(* IEC 61131-3 sources: guidance-for-physical-ai-production-designer-on-aws/source/plan2cell/examples/welding_cell_2_small/plc/trust/robot1/src, 20 files *)

(* ---- E_PlayerState.st ---- *)
(*
 * E_PlayerState
 * States of FB_ProgramPlayer (robot side of the bt2plc zone protocol).
 * Device simulator R1 (robot1), cell welding_cell_2_small. Generated by bt2plc 0.1.0.
 *)

TYPE E_PlayerState :
(
    PS_IDLE         := 0,    (* No program, pose held *)
    PS_NEXT_OP      := 10,   (* Advance to the next op: wStep := k, REQUEST := mask *)
    PS_WAIT_GRANT   := 20,   (* Wait (GRANT AND mask) = mask *)
    PS_DELAY        := 30,   (* Start delay of the op *)
    PS_MOVE         := 40,   (* Trajectory / blind home move *)
    PS_HOLD         := 50,   (* Hold at the end pose *)
    PS_WAIT_RELEASE := 60,   (* REQUEST := 0, wait (GRANT AND mask) = 0 *)
    PS_DONE         := 90,   (* Program finished *)
    PS_ERROR        := 99    (* Program aborted with an error *)
);
END_TYPE

(* ---- E_ProgramState.st ---- *)
(*
 * E_ProgramState
 * VW VASS standard - robot program states.
 * Device simulator R1 (robot1), cell welding_cell_2_small. Generated by bt2plc 0.1.0.
 *)

TYPE E_ProgramState :
(
    PRG_IDLE     := 0,
    PRG_RUNNING  := 1,
    PRG_STOPPED  := 2,
    PRG_PAUSED   := 3,
    PRG_FINISHED := 4,
    PRG_ERROR    := 5
);
END_TYPE

(* ---- E_RobotMode.st ---- *)
(*
 * E_RobotMode
 * VW VASS standard - KUKA KR C4 robot operating modes.
 * Device simulator R1 (robot1), cell welding_cell_2_small. Generated by bt2plc 0.1.0.
 *)

TYPE E_RobotMode :
(
    MODE_UNKNOWN := 0,
    MODE_T1      := 1,       (* Test mode 1 - reduced speed *)
    MODE_T2      := 2,       (* Test mode 2 - programmed speed *)
    MODE_AUT     := 3,       (* Automatic mode *)
    MODE_EXT     := 4        (* External automatic - PLC controlled *)
);
END_TYPE

(* ---- ST_OpDef.st ---- *)
(*
 * ST_OpDef
 * One op of the bt2plc robot program (row of GVL_Program.aOps).
 * Op k plays waypoints GVL_Program.aWp[nFirstWp..nLastWp] under the zone mask dwZoneMask.
 * Blind home op: bBlindHome = TRUE, nFirstWp = nLastWp = 0 (joint move to arHomeDeg over R_HOME_S).
 * Device simulator R1 (robot1), cell welding_cell_2_small. Generated by bt2plc 0.1.0.
 *)

TYPE ST_OpDef :
STRUCT
    sName           : STRING(32);   (* Operation id, e.g. 'W01' *)
    nFirstWp        : INT;          (* First waypoint index in aWp (0 = none) *)
    nLastWp         : INT;          (* Last waypoint index in aWp (0 = none) *)
    dwZoneMask      : DWORD;        (* REQUEST/GRANT bits (zones 0..30, bit 31 = permit) *)
    tDelay          : TIME;         (* Start delay after the grant *)
    tHold           : TIME;         (* Hold time at the end pose *)
    rDelay_s        : REAL;         (* Start delay in s (used by FB_ProgramPlayer) *)
    rHold_s         : REAL;         (* Hold time in s (used by FB_ProgramPlayer) *)
    rVelScale       : REAL;         (* Velocity scale of the trajectory (1.0 = nominal) *)
    bBlindHome      : BOOL;         (* TRUE = blind joint move to the home pose *)
END_STRUCT
END_TYPE

(* ---- ST_PROFIsafe_Trailer.st ---- *)
(*
 * ST_PROFIsafe_Trailer
 * PROFIsafe trailer - 4 bytes appended by the safety layer (status + 3-byte CRC).
 * Device simulator R1 (robot1), cell welding_cell_2_small. Generated by bt2plc 0.1.0.
 *)

TYPE ST_PROFIsafe_Trailer :
STRUCT
    byStatus        : BYTE;                     (* Status/Control byte *)
    abyCRC          : ARRAY[0..2] OF BYTE;      (* 3-byte CRC *)
END_STRUCT
END_TYPE

(* ---- ST_SafeInput.st ---- *)
(*
 * ST_SafeInput
 * PROFIsafe (Slot 1 - FDIO64) safe inputs: robot -> PLC, 8 bytes user data.
 * GSDML: 8x Unsigned8 Input + F_MessageTrailer4Byte.
 * Device simulator R1 (robot1), cell welding_cell_2_small. Generated by bt2plc 0.1.0.
 *)

TYPE ST_SafeInput :
STRUCT
    (* Byte 0: Safe robot status *)
    bSafe_DrivesOK          : BOOL;   (* Bit 0: Safe drives monitoring OK *)
    bSafe_RobotStopped      : BOOL;   (* Bit 1: Robot safely stopped (SOS/SS1) *)
    bSafe_ReducedSpeed      : BOOL;   (* Bit 2: Safe reduced speed active (SLS) *)
    bSafe_AxisMonitoring    : BOOL;   (* Bit 3: Safe axis range monitoring OK *)
    bSafe_ToolOK            : BOOL;   (* Bit 4: Safe tool monitoring OK *)
    bSafe_WorkspaceOK       : BOOL;   (* Bit 5: Safe workspace monitoring OK *)
    bSafe_Reserved06        : BOOL;   (* Bit 6: Reserved *)
    bSafe_Reserved07        : BOOL;   (* Bit 7: Reserved *)

    (* Byte 1: Safe gate/zone status *)
    bSafe_Gate1Closed       : BOOL;   (* Bit 0: Safety gate 1 closed *)
    bSafe_Gate2Closed       : BOOL;   (* Bit 1: Safety gate 2 closed *)
    bSafe_Gate3Closed       : BOOL;   (* Bit 2: Safety gate 3 closed *)
    bSafe_LightCurtainOK    : BOOL;   (* Bit 3: Light curtain free *)
    bSafe_EStopOK           : BOOL;   (* Bit 4: E-Stop not pressed (NC) *)
    bSafe_EnablingDevice    : BOOL;   (* Bit 5: Enabling device pressed (T1/T2) *)
    bSafe_OperatorSafe      : BOOL;   (* Bit 6: Operator protection OK *)
    bSafe_Reserved17        : BOOL;   (* Bit 7: Reserved *)

    (* Byte 2: Extended safe status *)
    bSafe_STO_Active        : BOOL;   (* Bit 0: Safe Torque Off active *)
    bSafe_SS1_Active        : BOOL;   (* Bit 1: Safe Stop 1 active *)
    bSafe_SS2_Active        : BOOL;   (* Bit 2: Safe Stop 2 active *)
    bSafe_SOS_Active        : BOOL;   (* Bit 3: Safe Operating Stop active *)
    bSafe_SLS_Active        : BOOL;   (* Bit 4: Safely-Limited Speed active *)
    bSafe_SLP_Active        : BOOL;   (* Bit 5: Safely-Limited Position active *)
    bSafe_Reserved26        : BOOL;   (* Bit 6: Reserved *)
    bSafe_FaultPresent      : BOOL;   (* Bit 7: Safety fault present *)

    (* Bytes 3-7: Additional safe signals *)
    bySafe_UserInput3       : BYTE;   (* Byte 3: User safe input *)
    bySafe_UserInput4       : BYTE;   (* Byte 4: User safe input *)
    bySafe_UserInput5       : BYTE;   (* Byte 5: User safe input *)
    bySafe_UserInput6       : BYTE;   (* Byte 6: User safe input *)
    bySafe_UserInput7       : BYTE;   (* Byte 7: User safe input *)
END_STRUCT
END_TYPE

(* ---- ST_SafeOutput.st ---- *)
(*
 * ST_SafeOutput
 * PROFIsafe (Slot 1 - FDIO64) safe outputs: PLC -> robot, 8 bytes user data.
 * GSDML: 8x Unsigned8 Output + F_MessageTrailer4Byte.
 * Device simulator R1 (robot1), cell welding_cell_2_small. Generated by bt2plc 0.1.0.
 *)

TYPE ST_SafeOutput :
STRUCT
    (* Byte 0: Safe control from PLC *)
    bSafe_DriveEnable       : BOOL;   (* Bit 0: Enable drives (safe channel) *)
    bSafe_ExternalEStop     : BOOL;   (* Bit 1: External E-Stop request *)
    bSafe_SafeStop1         : BOOL;   (* Bit 2: Request Safe Stop 1 *)
    bSafe_SafeStop2         : BOOL;   (* Bit 3: Request Safe Stop 2 *)
    bSafe_ReducedSpeedReq   : BOOL;   (* Bit 4: Request safe reduced speed *)
    bSafe_GateOverride      : BOOL;   (* Bit 5: Gate override (maintenance) *)
    bSafe_Reserved06        : BOOL;   (* Bit 6: Reserved *)
    bSafe_Reserved07        : BOOL;   (* Bit 7: Reserved *)

    (* Byte 1: Safe zone control *)
    bSafe_Zone1Enable       : BOOL;   (* Bit 0: Enable workspace zone 1 *)
    bSafe_Zone2Enable       : BOOL;   (* Bit 1: Enable workspace zone 2 *)
    bSafe_Zone3Enable       : BOOL;   (* Bit 2: Enable workspace zone 3 *)
    bSafe_Zone4Enable       : BOOL;   (* Bit 3: Enable workspace zone 4 *)
    bSafe_Reserved14        : BOOL;   (* Bit 4: Reserved *)
    bSafe_Reserved15        : BOOL;   (* Bit 5: Reserved *)
    bSafe_Reserved16        : BOOL;   (* Bit 6: Reserved *)
    bSafe_Reserved17        : BOOL;   (* Bit 7: Reserved *)

    (* Bytes 2-7: Additional safe control *)
    bySafe_UserOutput2      : BYTE;   (* Byte 2: User safe output *)
    bySafe_UserOutput3      : BYTE;   (* Byte 3: User safe output *)
    bySafe_UserOutput4      : BYTE;   (* Byte 4: User safe output *)
    bySafe_UserOutput5      : BYTE;   (* Byte 5: User safe output *)
    bySafe_UserOutput6      : BYTE;   (* Byte 6: User safe output *)
    bySafe_UserOutput7      : BYTE;   (* Byte 7: User safe output *)
END_STRUCT
END_TYPE

(* ---- ST_VASS_ControlWord.st ---- *)
(*
 * ST_VASS_ControlWord
 * VASS PLC control word - output bytes 0-1 (PLC -> robot), Slot 2 DIO256.
 * Device simulator R1 (robot1), cell welding_cell_2_small. Generated by bt2plc 0.1.0.
 *)

TYPE ST_VASS_ControlWord :
STRUCT
    (* Byte 0 *)
    bDrivesOn           : BOOL;   (* Bit 0: Enable drives *)
    bProgStart          : BOOL;   (* Bit 1: Start program *)
    bProgStop           : BOOL;   (* Bit 2: Stop program *)
    bProgCancel         : BOOL;   (* Bit 3: Cancel program *)
    bModeRequest        : BOOL;   (* Bit 4: Request EXT mode *)
    bReset              : BOOL;   (* Bit 5: Reset error *)
    bHomeRequest        : BOOL;   (* Bit 6: Move to home *)
    bConfirm            : BOOL;   (* Bit 7: Confirm/acknowledge *)

    (* Byte 1 *)
    bJobRequest         : BOOL;   (* Bit 8: New job request *)
    bGripperOpen        : BOOL;   (* Bit 9: Open gripper *)
    bGripperClose       : BOOL;   (* Bit 10: Close gripper *)
    bPeriphRelease      : BOOL;   (* Bit 11: Release peripheral *)
    bSpeedOverride      : BOOL;   (* Bit 12: Apply speed override *)
    bReserved13         : BOOL;   (* Bit 13: Reserved *)
    bReserved14         : BOOL;   (* Bit 14: Reserved *)
    bReserved15         : BOOL;   (* Bit 15: Reserved *)
END_STRUCT
END_TYPE

(* ---- ST_VASS_InputTelegram.st ---- *)
(*
 * ST_VASS_InputTelegram
 * Full VASS input telegram - 32 bytes (robot -> PLC), Slot 2 DIO256 inputs.
 * bt2plc use: bytes 4-5 wCurrentStep = op index (GVL_Program.STEP_BYTE),
 *             bytes 16-27 joint angles A1..A6 (FB_JointAngleEncoder),
 *             bytes 28-31 zone REQUEST DWORD LE (GVL_Program.REQ_BYTE).
 * Device simulator R1 (robot1), cell welding_cell_2_small. Generated by bt2plc 0.1.0.
 *)

TYPE ST_VASS_InputTelegram :
STRUCT
    stStatusWord        : ST_VASS_StatusWord;     (* Bytes 0-1:   Status word *)
    wActiveJobNr        : WORD;                   (* Bytes 2-3:   Active job number *)
    wCurrentStep        : WORD;                   (* Bytes 4-5:   Current program step *)
    wSpeedActual        : WORD;                   (* Bytes 6-7:   Actual speed % *)
    wActiveToolNr       : WORD;                   (* Bytes 8-9:   Active tool number *)
    wErrorCode          : WORD;                   (* Bytes 10-11: Active error code *)
    wWarningCode        : WORD;                   (* Bytes 12-13: Active warning code *)
    wPositionX          : INT;                    (* Bytes 14-15: Position X (0.1mm) *)
    wPositionY          : INT;                    (* Bytes 16-17: Position Y (0.1mm) *)
    wPositionZ          : INT;                    (* Bytes 18-19: Position Z (0.1mm) *)
    wUserWord10         : WORD;                   (* Bytes 20-21: User data *)
    wUserWord11         : WORD;                   (* Bytes 22-23: User data *)
    wUserWord12         : WORD;                   (* Bytes 24-25: User data *)
    wUserWord13         : WORD;                   (* Bytes 26-27: User data *)
    wUserWord14         : WORD;                   (* Bytes 28-29: User data *)
    wUserWord15         : WORD;                   (* Bytes 30-31: User data *)
END_STRUCT
END_TYPE

(* ---- ST_VASS_OutputTelegram.st ---- *)
(*
 * ST_VASS_OutputTelegram
 * Full VASS output telegram - 32 bytes (PLC -> robot), Slot 2 DIO256 outputs.
 * bt2plc use: bytes 4-5 PLAN_ID WORD LE during a production job (GVL_Program.PLAN_ID_BYTE),
 *             bytes 12-15 zone GRANT DWORD LE (GVL_Program.GRANT_BYTE).
 * Device simulator R1 (robot1), cell welding_cell_2_small. Generated by bt2plc 0.1.0.
 *)

TYPE ST_VASS_OutputTelegram :
STRUCT
    stControlWord       : ST_VASS_ControlWord;    (* Bytes 0-1:   Control word *)
    wJobNr              : WORD;                   (* Bytes 2-3:   Requested job number *)
    wParameter1         : WORD;                   (* Bytes 4-5:   Parameter 1 *)
    wParameter2         : WORD;                   (* Bytes 6-7:   Parameter 2 *)
    wSpeedOverride      : WORD;                   (* Bytes 8-9:   Speed override % *)
    wToolRequest        : WORD;                   (* Bytes 10-11: Tool change request *)
    wUserWord6          : WORD;                   (* Bytes 12-13: User command data *)
    wUserWord7          : WORD;                   (* Bytes 14-15: User command data *)
    wUserWord8          : WORD;                   (* Bytes 16-17: User command data *)
    wUserWord9          : WORD;                   (* Bytes 18-19: User command data *)
    wUserWord10         : WORD;                   (* Bytes 20-21: User command data *)
    wUserWord11         : WORD;                   (* Bytes 22-23: User command data *)
    wUserWord12         : WORD;                   (* Bytes 24-25: User command data *)
    wUserWord13         : WORD;                   (* Bytes 26-27: User command data *)
    wUserWord14         : WORD;                   (* Bytes 28-29: User command data *)
    wUserWord15         : WORD;                   (* Bytes 30-31: User command data *)
END_STRUCT
END_TYPE

(* ---- ST_VASS_StatusWord.st ---- *)
(*
 * ST_VASS_StatusWord
 * VASS robot status word - input bytes 0-1 (robot -> PLC), Slot 2 DIO256.
 * Device simulator R1 (robot1), cell welding_cell_2_small. Generated by bt2plc 0.1.0.
 *)

TYPE ST_VASS_StatusWord :
STRUCT
    (* Byte 0 *)
    bDrivesPowered      : BOOL;   (* Bit 0: Drives are powered on *)
    bProgRunning        : BOOL;   (* Bit 1: Program is running *)
    bAtHome             : BOOL;   (* Bit 2: Robot at home position *)
    bInPosition         : BOOL;   (* Bit 3: Robot in target position *)
    bModeExt            : BOOL;   (* Bit 4: External automatic mode active *)
    bReady              : BOOL;   (* Bit 5: Robot ready for command *)
    bError              : BOOL;   (* Bit 6: Error present *)
    bWarning            : BOOL;   (* Bit 7: Warning present *)

    (* Byte 1 *)
    bSafetyGateOK       : BOOL;   (* Bit 8: Safety gate closed *)
    bEStopNotActive     : BOOL;   (* Bit 9: E-Stop NOT active (NC logic) *)
    bProgFinished       : BOOL;   (* Bit 10: Program/job finished *)
    bJobAcknowledge     : BOOL;   (* Bit 11: Job number acknowledged *)
    bToolActive         : BOOL;   (* Bit 12: Tool/gripper active *)
    bPartPresent        : BOOL;   (* Bit 13: Part present in gripper *)
    bPeriphReady        : BOOL;   (* Bit 14: Peripheral devices ready *)
    bMaintRequired      : BOOL;   (* Bit 15: Maintenance required *)
END_STRUCT
END_TYPE

(* ---- ST_Waypoint.st ---- *)
(*
 * ST_Waypoint
 * One trajectory waypoint (row of GVL_Program.aWp). Flat fields for portability.
 * rT = seconds from op start; angles in degrees (KUKA A1..A6 after joint sign/offset mapping).
 * Device simulator R1 (robot1), cell welding_cell_2_small. Generated by bt2plc 0.1.0.
 *)

TYPE ST_Waypoint :
STRUCT
    rT              : REAL;         (* Time from op start (s) *)
    rA1             : REAL;         (* Axis 1 (deg) *)
    rA2             : REAL;         (* Axis 2 (deg) *)
    rA3             : REAL;         (* Axis 3 (deg) *)
    rA4             : REAL;         (* Axis 4 (deg) *)
    rA5             : REAL;         (* Axis 5 (deg) *)
    rA6             : REAL;         (* Axis 6 (deg) *)
END_STRUCT
END_TYPE

(* ---- GVL_DeviceParams.st ---- *)
NAMESPACE GVL_DeviceParams
(*
 * GVL_DeviceParams
 * PROFINET device identity parameters.
 * Device simulator R1 (robot1, station kuka-robi1), cell welding_cell_2_small. Generated by bt2plc 0.1.0.
 *
 * These parameters configure how the CODESYS PROFINET Device presents itself
 * on the network. They MUST match what the Siemens PLC expects (from the GSDML).
 *
 * In CODESYS, these are typically set via:
 *   1. The "PROFINET Device IEC Objects" tab in the device editor
 *   2. Or programmatically by writing to the device parameter structure
 *
 * The CODESYS PROFINET Device stack reads these at startup and uses them
 * in DCP responses and during the PROFINET connection establishment.
 *
 * IMPORTANT: The default CODESYS values (VendorId=0x02CC, DeviceId=0x1017)
 * will NOT work with the Siemens PLC that expects KUKA (0x019B / 0x0301).
 * You MUST override them.
 *)

{attribute 'qualified_only'}
VAR_GLOBAL
    (* === KUKA VKRCnexxt Device Identity === *)
    (* These values come from GSDML-V2.25-KUKA-Roboter-GmbH-VKR C4-Device-V1.0 *)

    VENDOR_ID           : UINT        := 16#019B;                 (* KUKA Roboter GmbH *)
    DEVICE_ID           : UINT        := 16#0301;                 (* VKR C4 Device *)
    STATION_TYPE        : STRING(240) := 'KUKA VKR C4';           (* Station type string *)
    DEVICE_TYPE         : STRING(28)  := 'KUKA VKR C4';           (* Device type string *)
    ORDER_ID            : STRING(20)  := 'KUKA VKRC nexxt';       (* Order number *)
    HW_REVISION         : UINT        := 1;                       (* Hardware revision *)
    SW_REV_PREFIX       : USINT       := 16#56;                   (* 'V' in ASCII *)
    SW_REV_MAJOR        : UINT        := 8;                       (* V8.x *)
    SW_REV_MINOR        : UINT        := 2;                       (* x.2 *)
    SW_REV_PATCH        : UINT        := 0;                       (* x.x.0 *)

    (* === Module Identification Numbers (from GSDML) === *)
    MODULE_IDENT_DAP    : DWORD       := DWORD#16#00000301;       (* DAP - Slot 0 *)
    MODULE_IDENT_FDIO64 : DWORD       := DWORD#16#0000008F;       (* PROFIsafe - Slot 1 *)
    MODULE_IDENT_DIO256 : DWORD       := DWORD#16#00001000;       (* VASS telegram - Slot 2 *)
    SUBMODULE_IDENT     : DWORD       := DWORD#16#00000001;       (* Submodule ident (all slots) *)

    (* === PROFIsafe Parameters (Slot 1) === *)
    (* These must match the F-parameter record in the PLC safety configuration *)
    F_SIL_LEVEL         : UINT        := 3;                       (* SIL 3 *)
    F_CRC_LENGTH        : UINT        := 3;                       (* 3-byte CRC *)
    F_WD_TIME_DEFAULT   : UINT        := 500;                     (* Watchdog 500ms *)
    F_BLOCK_ID          : UINT        := 0;                       (* Block ID *)
    F_PAR_CRC_DEFAULT   : UINT        := 16#FF59;                 (* Default F_Par_CRC = 65369 *)
END_VAR
END_NAMESPACE

(* ---- GVL_IO.st ---- *)
NAMESPACE GVL_IO
(*
 * GVL_IO
 * Global variable list for the PROFINET device I/O mapping.
 * Device simulator R1 (robot1, station kuka-robi1), cell welding_cell_2_small. Generated by bt2plc 0.1.0.
 *
 * These variables are mapped to the PROFINET device modules via the I/O Mapping tab.
 * Do NOT use AT addresses - the mapping is done in the device configuration.
 * Only PLC_PRG accesses this GVL: it copies the commands into local images and writes
 * the robot status back as a whole array / as scalars (the FBs never touch GVL_IO).
 *
 * Module mapping (set in I/O Mapping tab of each module):
 *   SafeIO_FDIO64 (Slot 1):
 *     "8 safe digital inputs" channels  -> GVL_IO.bySafeIn0..bySafeIn7
 *     "8 safe digital outputs" channels -> GVL_IO.bySafeOut0..bySafeOut7
 *
 *   VASS_DIO256 (Slot 2):
 *     Input channel  -> GVL_IO.aVassInputData
 *     Output channel -> GVL_IO.aVassOutputData
 *)

{attribute 'qualified_only'}
VAR_GLOBAL
    (* ========================================================================
       SLOT 1 - PROFIsafe FDIO64 Module
       8 individual USINT/BYTE channels per direction
       Map each one to the corresponding "8 safe digital inputs/outputs" row
       ======================================================================== *)

    (* Safe Inputs: Robot -> PLC (mapped to "8 safe digital inputs" channels) *)
    bySafeIn0       : BYTE;     (* Safe input byte 0: Drive status *)
    bySafeIn1       : BYTE;     (* Safe input byte 1: Gate/protection *)
    bySafeIn2       : BYTE;     (* Safe input byte 2: STO/SS1/SS2/SOS/SLS *)
    bySafeIn3       : BYTE;     (* Safe input byte 3: User *)
    bySafeIn4       : BYTE;     (* Safe input byte 4: User *)
    bySafeIn5       : BYTE;     (* Safe input byte 5: User *)
    bySafeIn6       : BYTE;     (* Safe input byte 6: User *)
    bySafeIn7       : BYTE;     (* Safe input byte 7: User *)

    (* Safe Outputs: PLC -> Robot (mapped to "8 safe digital outputs" channels) *)
    bySafeOut0      : BYTE;     (* Safe output byte 0: Drive enable, E-Stop, SS1/SS2 *)
    bySafeOut1      : BYTE;     (* Safe output byte 1: Zone enables *)
    bySafeOut2      : BYTE;     (* Safe output byte 2: User *)
    bySafeOut3      : BYTE;     (* Safe output byte 3: User *)
    bySafeOut4      : BYTE;     (* Safe output byte 4: User *)
    bySafeOut5      : BYTE;     (* Safe output byte 5: User *)
    bySafeOut6      : BYTE;     (* Safe output byte 6: User *)
    bySafeOut7      : BYTE;     (* Safe output byte 7: User *)

    (* ========================================================================
       SLOT 2 - DIO256 VASS Telegram
       32 bytes per direction as arrays
       ======================================================================== *)

    (* VASS Inputs: Robot -> PLC (32 bytes) *)
    aVassInputData      : ARRAY[0..31] OF BYTE;

    (* VASS Outputs: PLC -> Robot (32 bytes) *)
    aVassOutputData     : ARRAY[0..31] OF BYTE;
END_VAR
END_NAMESPACE

(* ---- GVL_Program.st ---- *)
NAMESPACE GVL_Program
(*
 * GVL_Program - generated by bt2plc 0.1.0 - DO NOT EDIT
 * Robot program of robot1 (R1) for plan bt_1790934549_welding_cell_2_small (cell welding_cell_2_small)
 * Angles in degrees (KUKA A1..A6 after joint sign/offset), times in seconds from op start.
 *)
{attribute 'qualified_only'}
VAR_GLOBAL
    (* ========================================================================
       IDENTITY / PROTOCOL
       ======================================================================== *)
    ROBOT_TAG               : STRING(16) := 'R1';
    ROBOT_NS                : STRING(32) := 'robot1';
    ROBOT_INDEX             : WORD := WORD#1;
    PLAN_ID                 : WORD := WORD#16#F77E;             (* must match the head PLC *)
    PROD_FOLGE              : WORD := WORD#11;
    HOME_FOLGE              : WORD := WORD#125;
    JOB_NUMBER_BYTE         : BOOL := FALSE;
    STEP_BYTE               : INT := 4;
    REQ_BYTE                : INT := 28;
    GRANT_BYTE              : INT := 12;
    PLAN_ID_BYTE            : INT := 4;
    R_TASK_S                : REAL := 0.0200;                   (* device MainTask interval *)
    R_HOME_S                : REAL := 7.0000;                   (* blind home duration *)
    R_AT_HOME_TOL_DEG       : REAL := 0.5000;
    R_START_TOL_DEG         : REAL := 1.0000;
    ERR_UNKNOWN_FOLGE       : WORD := WORD#16#0101;
    ERR_PLAN_MISMATCH       : WORD := WORD#16#0103;
    WARN_START_DEVIATION    : WORD := WORD#16#0201;

    (* ========================================================================
       PROGRAM
       ======================================================================== *)
    N_OPS                   : INT := 8;
    N_WP                    : INT := 211;
    arHomeDeg               : ARRAY[1..6] OF REAL := [0.0000, -90.0000, 90.0000, 0.0000, 0.0000, 0.0000];
    aOps                    : ARRAY[1..8] OF ST_OpDef := [
        (sName := 'W01', nFirstWp := 1, nLastWp := 47, dwZoneMask := DWORD#16#00000001, tDelay := T#0MS, tHold := T#500MS, rDelay_s := 0.0000, rHold_s := 0.5000, rVelScale := 1.0000, bBlindHome := FALSE),    (* #1 W01 (weld) *)
        (sName := 'W02', nFirstWp := 48, nLastWp := 68, dwZoneMask := DWORD#16#00000002, tDelay := T#0MS, tHold := T#500MS, rDelay_s := 0.0000, rHold_s := 0.5000, rVelScale := 1.0000, bBlindHome := FALSE),    (* #2 W02 (weld) *)
        (sName := 'W03', nFirstWp := 69, nLastWp := 95, dwZoneMask := DWORD#16#00000001, tDelay := T#0MS, tHold := T#500MS, rDelay_s := 0.0000, rHold_s := 0.5000, rVelScale := 1.0000, bBlindHome := FALSE),    (* #3 W03 (weld) *)
        (sName := 'W06', nFirstWp := 96, nLastWp := 110, dwZoneMask := DWORD#16#00000002, tDelay := T#0MS, tHold := T#500MS, rDelay_s := 0.0000, rHold_s := 0.5000, rVelScale := 1.0000, bBlindHome := FALSE),    (* #4 W06 (weld) *)
        (sName := 'W05', nFirstWp := 111, nLastWp := 137, dwZoneMask := DWORD#16#00000001, tDelay := T#0MS, tHold := T#500MS, rDelay_s := 0.0000, rHold_s := 0.5000, rVelScale := 1.0000, bBlindHome := FALSE),    (* #5 W05 (weld) *)
        (sName := 'W04', nFirstWp := 138, nLastWp := 159, dwZoneMask := DWORD#16#00000002, tDelay := T#0MS, tHold := T#500MS, rDelay_s := 0.0000, rHold_s := 0.5000, rVelScale := 1.0000, bBlindHome := FALSE),    (* #6 W04 (weld) *)
        (sName := 'R1_PARK', nFirstWp := 160, nLastWp := 169, dwZoneMask := DWORD#16#00000001, tDelay := T#0MS, tHold := T#500MS, rDelay_s := 0.0000, rHold_s := 0.5000, rVelScale := 1.0000, bBlindHome := FALSE),    (* #7 R1_PARK (move) *)
        (sName := 'HOME', nFirstWp := 170, nLastWp := 211, dwZoneMask := DWORD#16#00000002, tDelay := T#0MS, tHold := T#0MS, rDelay_s := 0.0000, rHold_s := 0.0000, rVelScale := 1.0000, bBlindHome := FALSE)    (* #8 HOME (home) *)
    ];
    aWp                     : ARRAY[1..211] OF ST_Waypoint := [
        (* op 1 W01 - traj_robot1_W01 *)
        (rT := 0.0000, rA1 := 0.0000, rA2 := -90.0000, rA3 := 90.0000, rA4 := 0.0000, rA5 := 0.0000, rA6 := 0.0000),
        (rT := 0.2677, rA1 := -0.2925, rA2 := -89.9560, rA3 := 90.0355, rA4 := 0.0753, rA5 := 0.1975, rA6 := 0.0896),
        (rT := 0.5350, rA1 := -1.1481, rA2 := -89.8273, rA3 := 90.1392, rA4 := 0.2955, rA5 := 0.7752, rA6 := 0.3515),
        (rT := 0.8027, rA1 := -2.5335, rA2 := -89.6188, rA3 := 90.3072, rA4 := 0.6521, rA5 := 1.7108, rA6 := 0.7756),
        (rT := 1.0703, rA1 := -4.4157, rA2 := -89.3356, rA3 := 90.5354, rA4 := 1.1366, rA5 := 2.9817, rA6 := 1.3518),
        (rT := 1.3377, rA1 := -6.7615, rA2 := -88.9827, rA3 := 90.8198, rA4 := 1.7404, rA5 := 4.5657, rA6 := 2.0699),
        (rT := 1.6053, rA1 := -9.5379, rA2 := -88.5650, rA3 := 91.1564, rA4 := 2.4550, rA5 := 6.4405, rA6 := 2.9199),
        (rT := 1.8730, rA1 := -12.7117, rA2 := -88.0875, rA3 := 91.5412, rA4 := 3.2720, rA5 := 8.5836, rA6 := 3.8915),
        (rT := 2.1403, rA1 := -16.2497, rA2 := -87.5551, rA3 := 91.9702, rA4 := 4.1827, rA5 := 10.9727, rA6 := 4.9746),
        (rT := 2.4080, rA1 := -20.1190, rA2 := -86.9730, rA3 := 92.4393, rA4 := 5.1786, rA5 := 13.5854, rA6 := 6.1591),
        (rT := 2.6757, rA1 := -24.2863, rA2 := -86.3460, rA3 := 92.9446, rA4 := 6.2512, rA5 := 16.3994, rA6 := 7.4349),
        (rT := 2.9430, rA1 := -28.7185, rA2 := -85.6792, rA3 := 93.4820, rA4 := 7.3921, rA5 := 19.3923, rA6 := 8.7918),
        (rT := 3.2107, rA1 := -33.3826, rA2 := -84.9774, rA3 := 94.0475, rA4 := 8.5926, rA5 := 22.5417, rA6 := 10.2196),
        (rT := 3.4783, rA1 := -38.2454, rA2 := -84.2458, rA3 := 94.6371, rA4 := 9.8443, rA5 := 25.8253, rA6 := 11.7083),
        (rT := 3.7457, rA1 := -43.2738, rA2 := -83.4892, rA3 := 95.2467, rA4 := 11.1386, rA5 := 29.2207, rA6 := 13.2477),
        (rT := 4.0133, rA1 := -48.4346, rA2 := -82.7128, rA3 := 95.8725, rA4 := 12.4670, rA5 := 32.7056, rA6 := 14.8276),
        (rT := 4.2810, rA1 := -53.6948, rA2 := -81.9214, rA3 := 96.5102, rA4 := 13.8209, rA5 := 36.2575, rA6 := 16.4379),
        (rT := 4.5483, rA1 := -59.0212, rA2 := -81.1200, rA3 := 97.1561, rA4 := 15.1919, rA5 := 39.8542, rA6 := 18.0685),
        (rT := 4.8160, rA1 := -64.3808, rA2 := -80.3136, rA3 := 97.8059, rA4 := 16.5715, rA5 := 43.4732, rA6 := 19.7093),
        (rT := 5.0837, rA1 := -69.7403, rA2 := -79.5072, rA3 := 98.4557, rA4 := 17.9510, rA5 := 47.0923, rA6 := 21.3500),
        (rT := 5.3510, rA1 := -75.0667, rA2 := -78.7058, rA3 := 99.1015, rA4 := 19.3220, rA5 := 50.6890, rA6 := 22.9806),
        (rT := 5.6187, rA1 := -80.3269, rA2 := -77.9144, rA3 := 99.7393, rA4 := 20.6760, rA5 := 54.2409, rA6 := 24.5910),
        (rT := 5.8863, rA1 := -85.4878, rA2 := -77.1379, rA3 := 100.3650, rA4 := 22.0044, rA5 := 57.7258, rA6 := 26.1709),
        (rT := 6.1537, rA1 := -90.5161, rA2 := -76.3814, rA3 := 100.9747, rA4 := 23.2987, rA5 := 61.1212, rA6 := 27.7103),
        (rT := 6.4213, rA1 := -95.3789, rA2 := -75.6498, rA3 := 101.5643, rA4 := 24.5503, rA5 := 64.4048, rA6 := 29.1989),
        (rT := 6.6890, rA1 := -100.0430, rA2 := -74.9480, rA3 := 102.1298, rA4 := 25.7509, rA5 := 67.5542, rA6 := 30.6268),
        (rT := 6.9563, rA1 := -104.4752, rA2 := -74.2812, rA3 := 102.6671, rA4 := 26.8917, rA5 := 70.5471, rA6 := 31.9836),
        (rT := 7.2240, rA1 := -108.6425, rA2 := -73.6542, rA3 := 103.1724, rA4 := 27.9644, rA5 := 73.3611, rA6 := 33.2594),
        (rT := 7.4917, rA1 := -112.5118, rA2 := -73.0720, rA3 := 103.6415, rA4 := 28.9603, rA5 := 75.9738, rA6 := 34.4439),
        (rT := 7.7590, rA1 := -116.0498, rA2 := -72.5397, rA3 := 104.0705, rA4 := 29.8710, rA5 := 78.3629, rA6 := 35.5271),
        (rT := 8.0267, rA1 := -119.2236, rA2 := -72.0622, rA3 := 104.4553, rA4 := 30.6879, rA5 := 80.5060, rA6 := 36.4987),
        (rT := 8.2943, rA1 := -122.0000, rA2 := -71.6445, rA3 := 104.7919, rA4 := 31.4026, rA5 := 82.3807, rA6 := 37.3486),
        (rT := 8.5617, rA1 := -124.3458, rA2 := -71.2916, rA3 := 105.0764, rA4 := 32.0064, rA5 := 83.9648, rA6 := 38.0668),
        (rT := 8.8293, rA1 := -126.2280, rA2 := -71.0084, rA3 := 105.3046, rA4 := 32.4908, rA5 := 85.2357, rA6 := 38.6430),
        (rT := 9.0970, rA1 := -127.6134, rA2 := -70.7999, rA3 := 105.4725, rA4 := 32.8474, rA5 := 86.1712, rA6 := 39.0671),
        (rT := 9.3643, rA1 := -128.4690, rA2 := -70.6712, rA3 := 105.5763, rA4 := 33.0677, rA5 := 86.7489, rA6 := 39.3290),
        (rT := 9.6320, rA1 := -128.7615, rA2 := -70.6272, rA3 := 105.6117, rA4 := 33.1430, rA5 := 86.9465, rA6 := 39.4186),
        (rT := 9.7320, rA1 := -128.7615, rA2 := -70.2228, rA3 := 105.9156, rA4 := 33.1800, rA5 := 86.8872, rA6 := 39.3731),
        (rT := 9.8320, rA1 := -128.7615, rA2 := -69.6268, rA3 := 106.3586, rA4 := 33.2522, rA5 := 86.7080, rA6 := 39.2426),
        (rT := 9.9320, rA1 := -128.7615, rA2 := -69.3317, rA3 := 106.5670, rA4 := 33.3382, rA5 := 86.3784, rA6 := 39.0108),
        (rT := 10.0320, rA1 := -128.7615, rA2 := -69.0945, rA3 := 106.7257, rA4 := 33.4236, rA5 := 85.9874, rA6 := 38.7386),
        (rT := 10.1320, rA1 := -128.7615, rA2 := -68.8270, rA3 := 106.9027, rA4 := 33.4818, rA5 := 85.6233, rA6 := 38.4888),
        (rT := 10.2320, rA1 := -128.7615, rA2 := -68.5576, rA3 := 107.0760, rA4 := 33.5282, rA5 := 85.2576, rA6 := 38.2401),
        (rT := 10.3320, rA1 := -128.7615, rA2 := -68.2851, rA3 := 107.2465, rA4 := 33.5686, rA5 := 84.8912, rA6 := 37.9919),
        (rT := 10.4320, rA1 := -128.7615, rA2 := -68.0100, rA3 := 107.4140, rA4 := 33.6041, rA5 := 84.5242, rA6 := 37.7441),
        (rT := 10.5320, rA1 := -128.7615, rA2 := -67.6617, rA3 := 107.6183, rA4 := 33.6457, rA5 := 84.0653, rA6 := 37.4348),
        (rT := 10.6320, rA1 := -128.7615, rA2 := -67.4517, rA3 := 107.7396, rA4 := 33.6697, rA5 := 83.7898, rA6 := 37.2493),
        (* op 2 W02 - traj_robot1_W02 *)
        (rT := 0.0000, rA1 := -128.7615, rA2 := -67.4517, rA3 := 107.7396, rA4 := 33.6697, rA5 := 83.7898, rA6 := 37.2493),
        (rT := 0.2820, rA1 := -128.6426, rA2 := -67.6366, rA3 := 107.8186, rA4 := 32.7502, rA5 := 82.9536, rA6 := 37.7433),
        (rT := 0.5643, rA1 := -128.3199, rA2 := -68.1386, rA3 := 108.0329, rA4 := 30.2544, rA5 := 80.6837, rA6 := 39.0840),
        (rT := 0.8463, rA1 := -127.8443, rA2 := -68.8784, rA3 := 108.3488, rA4 := 26.5764, rA5 := 77.3387, rA6 := 41.0597),
        (rT := 1.1283, rA1 := -127.2668, rA2 := -69.7767, rA3 := 108.7324, rA4 := 22.1103, rA5 := 73.2769, rA6 := 43.4588),
        (rT := 1.4103, rA1 := -126.6384, rA2 := -70.7542, rA3 := 109.1498, rA4 := 17.2501, rA5 := 68.8567, rA6 := 46.0696),
        (rT := 1.6927, rA1 := -126.0100, rA2 := -71.7318, rA3 := 109.5672, rA4 := 12.3899, rA5 := 64.4365, rA6 := 48.6804),
        (rT := 1.9747, rA1 := -125.4325, rA2 := -72.6301, rA3 := 109.9508, rA4 := 7.9238, rA5 := 60.3747, rA6 := 51.0796),
        (rT := 2.2567, rA1 := -124.9570, rA2 := -73.3699, rA3 := 110.2667, rA4 := 4.2458, rA5 := 57.0297, rA6 := 53.0553),
        (rT := 2.5390, rA1 := -124.6342, rA2 := -73.8718, rA3 := 110.4810, rA4 := 1.7500, rA5 := 54.7598, rA6 := 54.3960),
        (rT := 2.8210, rA1 := -124.5154, rA2 := -74.0568, rA3 := 110.5600, rA4 := 0.8305, rA5 := 53.9236, rA6 := 54.8899),
        (rT := 2.9210, rA1 := -124.5151, rA2 := -73.6213, rA3 := 110.8768, rA4 := 0.5687, rA5 := 53.3206, rA6 := 55.0767),
        (rT := 3.0210, rA1 := -124.5148, rA2 := -72.9810, rA3 := 111.3378, rA4 := 0.2163, rA5 := 52.4162, rA6 := 55.3282),
        (rT := 3.1210, rA1 := -124.5148, rA2 := -72.6684, rA3 := 111.5513, rA4 := 0.1257, rA5 := 51.9277, rA6 := 55.3932),
        (rT := 3.2210, rA1 := -124.5148, rA2 := -72.4184, rA3 := 111.7128, rA4 := 0.1050, rA5 := 51.5125, rA6 := 55.4084),
        (rT := 3.3210, rA1 := -124.5148, rA2 := -72.1325, rA3 := 111.8956, rA4 := 0.0727, rA5 := 51.0535, rA6 := 55.4318),
        (rT := 3.4210, rA1 := -124.5148, rA2 := -71.8436, rA3 := 112.0754, rA4 := 0.0510, rA5 := 50.5913, rA6 := 55.4476),
        (rT := 3.5210, rA1 := -124.5148, rA2 := -71.5517, rA3 := 112.2520, rA4 := 0.0354, rA5 := 50.1273, rA6 := 55.4590),
        (rT := 3.6210, rA1 := -124.5148, rA2 := -71.2569, rA3 := 112.4255, rA4 := 0.0248, rA5 := 49.6619, rA6 := 55.4668),
        (rT := 3.7210, rA1 := -124.5148, rA2 := -70.8835, rA3 := 112.6373, rA4 := 0.0160, rA5 := 49.0790, rA6 := 55.4732),
        (rT := 3.8210, rA1 := -124.5148, rA2 := -70.6583, rA3 := 112.7632, rA4 := 0.0121, rA5 := 48.7290, rA6 := 55.4761),
        (* op 3 W03 - traj_robot1_W03 *)
        (rT := 0.0000, rA1 := -124.5148, rA2 := -70.6583, rA3 := 112.7632, rA4 := 0.0121, rA5 := 48.7290, rA6 := 55.4761),
        (rT := 0.2767, rA1 := -124.4617, rA2 := -70.7313, rA3 := 112.7862, rA4 := -0.6572, rA5 := 48.6812, rA6 := 55.9965),
        (rT := 0.5530, rA1 := -124.3117, rA2 := -70.9378, rA3 := 112.8512, rA4 := -2.5487, rA5 := 48.5461, rA6 := 57.4671),
        (rT := 0.8297, rA1 := -124.0786, rA2 := -71.2585, rA3 := 112.9524, rA4 := -5.4877, rA5 := 48.3361, rA6 := 59.7523),
        (rT := 1.1063, rA1 := -123.7762, rA2 := -71.6746, rA3 := 113.0835, rA4 := -9.2998, rA5 := 48.0639, rA6 := 62.7161),
        (rT := 1.3830, rA1 := -123.4185, rA2 := -72.1669, rA3 := 113.2386, rA4 := -13.8102, rA5 := 47.7417, rA6 := 66.2230),
        (rT := 1.6593, rA1 := -123.0192, rA2 := -72.7163, rA3 := 113.4118, rA4 := -18.8444, rA5 := 47.3821, rA6 := 70.1371),
        (rT := 1.9360, rA1 := -122.5922, rA2 := -73.3038, rA3 := 113.5970, rA4 := -24.2279, rA5 := 46.9976, rA6 := 74.3228),
        (rT := 2.2127, rA1 := -122.1513, rA2 := -73.9104, rA3 := 113.7882, rA4 := -29.7859, rA5 := 46.6006, rA6 := 78.6441),
        (rT := 2.4893, rA1 := -121.7105, rA2 := -74.5170, rA3 := 113.9794, rA4 := -35.3439, rA5 := 46.2036, rA6 := 82.9655),
        (rT := 2.7657, rA1 := -121.2835, rA2 := -75.1045, rA3 := 114.1646, rA4 := -40.7273, rA5 := 45.8191, rA6 := 87.1511),
        (rT := 3.0423, rA1 := -120.8842, rA2 := -75.6540, rA3 := 114.3378, rA4 := -45.7616, rA5 := 45.4595, rA6 := 91.0652),
        (rT := 3.3190, rA1 := -120.5264, rA2 := -76.1462, rA3 := 114.4929, rA4 := -50.2720, rA5 := 45.1373, rA6 := 94.5721),
        (rT := 3.5953, rA1 := -120.2241, rA2 := -76.5623, rA3 := 114.6241, rA4 := -54.0840, rA5 := 44.8650, rA6 := 97.5360),
        (rT := 3.8720, rA1 := -119.9910, rA2 := -76.8830, rA3 := 114.7252, rA4 := -57.0231, rA5 := 44.6551, rA6 := 99.8211),
        (rT := 4.1487, rA1 := -119.8409, rA2 := -77.0895, rA3 := 114.7902, rA4 := -58.9146, rA5 := 44.5200, rA6 := 101.2917),
        (rT := 4.4253, rA1 := -119.7879, rA2 := -77.1625, rA3 := 114.8133, rA4 := -59.5839, rA5 := 44.4722, rA6 := 101.8121),
        (rT := 4.5377, rA1 := -119.7876, rA2 := -76.7001, rA3 := 115.1416, rA4 := -60.3559, rA5 := 44.3240, rA6 := 102.6809),
        (rT := 4.6505, rA1 := -119.7872, rA2 := -76.0201, rA3 := 115.6192, rA4 := -61.4852, rA5 := 44.0795, rA6 := 103.9753),
        (rT := 4.7505, rA1 := -119.7872, rA2 := -75.6879, rA3 := 115.8405, rA4 := -62.0177, rA5 := 43.8942, rA6 := 104.6450),
        (rT := 4.8505, rA1 := -119.7872, rA2 := -75.4218, rA3 := 116.0082, rA4 := -62.4422, rA5 := 43.7024, rA6 := 105.2177),
        (rT := 4.9505, rA1 := -119.7872, rA2 := -75.1169, rA3 := 116.1984, rA4 := -62.9641, rA5 := 43.4812, rA6 := 105.9117),
        (rT := 5.0505, rA1 := -119.7872, rA2 := -74.8088, rA3 := 116.3854, rA4 := -63.4806, rA5 := 43.2578, rA6 := 106.6047),
        (rT := 5.1505, rA1 := -119.7872, rA2 := -74.4987, rA3 := 116.5684, rA4 := -63.9374, rA5 := 43.0597, rA6 := 107.2204),
        (rT := 5.2505, rA1 := -119.7872, rA2 := -74.1853, rA3 := 116.7483, rA4 := -64.3947, rA5 := 42.8625, rA6 := 107.8387),
        (rT := 5.3505, rA1 := -119.7872, rA2 := -73.7867, rA3 := 116.9688, rA4 := -65.0379, rA5 := 42.5916, rA6 := 108.7077),
        (rT := 5.4505, rA1 := -119.7872, rA2 := -73.5459, rA3 := 117.1000, rA4 := -65.4365, rA5 := 42.4249, rA6 := 109.2463),
        (* op 4 W06 - traj_robot1_W06 *)
        (rT := 0.0000, rA1 := -119.7872, rA2 := -73.5459, rA3 := 117.1000, rA4 := -65.4365, rA5 := 42.4249, rA6 := 109.2463),
        (rT := 0.2930, rA1 := -119.1489, rA2 := -72.8001, rA3 := 114.8711, rA4 := -64.2164, rA5 := 43.4199, rA6 := 108.0229),
        (rT := 0.5860, rA1 := -117.7444, rA2 := -71.1593, rA3 := 109.9675, rA4 := -61.5322, rA5 := 45.6090, rA6 := 105.3312),
        (rT := 0.8790, rA1 := -116.3400, rA2 := -69.5185, rA3 := 105.0638, rA4 := -58.8479, rA5 := 47.7981, rA6 := 102.6395),
        (rT := 1.1720, rA1 := -115.7016, rA2 := -68.7727, rA3 := 102.8349, rA4 := -57.6278, rA5 := 48.7931, rA6 := 101.4160),
        (rT := 1.2720, rA1 := -115.7012, rA2 := -68.3831, rA3 := 103.1319, rA4 := -57.6419, rA5 := 48.7925, rA6 := 101.4570),
        (rT := 1.3720, rA1 := -115.7007, rA2 := -67.8085, rA3 := 103.5655, rA4 := -57.7461, rA5 := 48.7415, rA6 := 101.6606),
        (rT := 1.4720, rA1 := -115.7006, rA2 := -67.5229, rA3 := 103.7711, rA4 := -58.0189, rA5 := 48.5849, rA6 := 102.1462),
        (rT := 1.5720, rA1 := -115.7007, rA2 := -67.2934, rA3 := 103.9284, rA4 := -58.3483, rA5 := 48.3900, rA6 := 102.7163),
        (rT := 1.6720, rA1 := -115.7007, rA2 := -67.0361, rA3 := 104.1022, rA4 := -58.6282, rA5 := 48.2163, rA6 := 103.1755),
        (rT := 1.7720, rA1 := -115.7007, rA2 := -66.7771, rA3 := 104.2724, rA4 := -58.9197, rA5 := 48.0319, rA6 := 103.6366),
        (rT := 1.8720, rA1 := -115.7007, rA2 := -66.5140, rA3 := 104.4406, rA4 := -59.2591, rA5 := 47.8179, rA6 := 104.1645),
        (rT := 1.9720, rA1 := -115.7007, rA2 := -66.2481, rA3 := 104.6058, rA4 := -59.6142, rA5 := 47.5951, rA6 := 104.7081),
        (rT := 2.0720, rA1 := -115.7007, rA2 := -65.9124, rA3 := 104.8068, rA4 := -60.0493, rA5 := 47.3267, rA6 := 105.3635),
        (rT := 2.1720, rA1 := -115.7007, rA2 := -65.7101, rA3 := 104.9261, rA4 := -60.3105, rA5 := 47.1665, rA6 := 105.7542),
        (* op 5 W05 - traj_robot1_W05 *)
        (rT := 0.0000, rA1 := -115.7007, rA2 := -65.7101, rA3 := 104.9261, rA4 := -60.3105, rA5 := 47.1665, rA6 := 105.7542),
        (rT := 0.2757, rA1 := -115.7494, rA2 := -65.7146, rA3 := 104.8564, rA4 := -59.6416, rA5 := 47.2762, rA6 := 105.2455),
        (rT := 0.5517, rA1 := -115.8870, rA2 := -65.7270, rA3 := 104.6592, rA4 := -57.7513, rA5 := 47.5859, rA6 := 103.8079),
        (rT := 0.8273, rA1 := -116.1007, rA2 := -65.7464, rA3 := 104.3529, rA4 := -54.8140, rA5 := 48.0672, rA6 := 101.5740),
        (rT := 1.1030, rA1 := -116.3780, rA2 := -65.7715, rA3 := 103.9556, rA4 := -51.0043, rA5 := 48.6915, rA6 := 98.6766),
        (rT := 1.3787, rA1 := -116.7061, rA2 := -65.8013, rA3 := 103.4855, rA4 := -46.4967, rA5 := 49.4301, rA6 := 95.2484),
        (rT := 1.6547, rA1 := -117.0722, rA2 := -65.8345, rA3 := 102.9609, rA4 := -41.4655, rA5 := 50.2545, rA6 := 91.4221),
        (rT := 1.9303, rA1 := -117.4638, rA2 := -65.8700, rA3 := 102.3998, rA4 := -36.0854, rA5 := 51.1361, rA6 := 87.3303),
        (rT := 2.2060, rA1 := -117.8681, rA2 := -65.9066, rA3 := 101.8205, rA4 := -30.5308, rA5 := 52.0463, rA6 := 83.1058),
        (rT := 2.4820, rA1 := -118.2723, rA2 := -65.9433, rA3 := 101.2413, rA4 := -24.9762, rA5 := 52.9565, rA6 := 78.8814),
        (rT := 2.7577, rA1 := -118.6639, rA2 := -65.9788, rA3 := 100.6802, rA4 := -19.5961, rA5 := 53.8381, rA6 := 74.7896),
        (rT := 3.0333, rA1 := -119.0301, rA2 := -66.0120, rA3 := 100.1555, rA4 := -14.5649, rA5 := 54.6625, rA6 := 70.9633),
        (rT := 3.3093, rA1 := -119.3582, rA2 := -66.0417, rA3 := 99.6854, rA4 := -10.0572, rA5 := 55.4012, rA6 := 67.5351),
        (rT := 3.5850, rA1 := -119.6354, rA2 := -66.0668, rA3 := 99.2881, rA4 := -6.2475, rA5 := 56.0254, rA6 := 64.6377),
        (rT := 3.8607, rA1 := -119.8492, rA2 := -66.0862, rA3 := 98.9818, rA4 := -3.3103, rA5 := 56.5068, rA6 := 62.4038),
        (rT := 4.1363, rA1 := -119.9868, rA2 := -66.0987, rA3 := 98.7847, rA4 := -1.4200, rA5 := 56.8165, rA6 := 60.9662),
        (rT := 4.4123, rA1 := -120.0355, rA2 := -66.1031, rA3 := 98.7149, rA4 := -0.7511, rA5 := 56.9261, rA6 := 60.4575),
        (rT := 4.5123, rA1 := -120.0357, rA2 := -65.7312, rA3 := 99.0104, rA4 := -0.6308, rA5 := 56.7548, rA6 := 60.3791),
        (rT := 4.6123, rA1 := -120.0360, rA2 := -65.1841, rA3 := 99.4405, rA4 := -0.4466, rA5 := 56.4312, rA6 := 60.2589),
        (rT := 4.7123, rA1 := -120.0360, rA2 := -64.9162, rA3 := 99.6405, rA4 := -0.3319, rA5 := 56.0924, rA6 := 60.1840),
        (rT := 4.8123, rA1 := -120.0359, rA2 := -64.7015, rA3 := 99.7923, rA4 := -0.2398, rA5 := 55.7079, rA6 := 60.1236),
        (rT := 4.9123, rA1 := -120.0359, rA2 := -64.4565, rA3 := 99.9636, rA4 := -0.1684, rA5 := 55.2797, rA6 := 60.0766),
        (rT := 5.0123, rA1 := -120.0359, rA2 := -64.2094, rA3 := 100.1316, rA4 := -0.1162, rA5 := 54.8474, rA6 := 60.0420),
        (rT := 5.1123, rA1 := -120.0359, rA2 := -63.9609, rA3 := 100.2959, rA4 := -0.0836, rA5 := 54.4700, rA6 := 60.0204),
        (rT := 5.2123, rA1 := -120.0359, rA2 := -63.7100, rA3 := 100.4571, rA4 := -0.0624, rA5 := 54.0904, rA6 := 60.0063),
        (rT := 5.3123, rA1 := -120.0359, rA2 := -63.3911, rA3 := 100.6546, rA4 := -0.0410, rA5 := 53.5493, rA6 := 59.9919),
        (rT := 5.4123, rA1 := -120.0359, rA2 := -63.1985, rA3 := 100.7720, rA4 := -0.0303, rA5 := 53.2125, rA6 := 59.9847),
        (* op 6 W04 - traj_robot1_W04 *)
        (rT := 0.0000, rA1 := -120.0359, rA2 := -63.1985, rA3 := 100.7720, rA4 := -0.0303, rA5 := 53.2125, rA6 := 59.9847),
        (rT := 0.2773, rA1 := -120.1288, rA2 := -63.1954, rA3 := 100.6111, rA4 := 0.7952, rA5 := 54.0248, rA6 := 59.6456),
        (rT := 0.5547, rA1 := -120.3834, rA2 := -63.1866, rA3 := 100.1699, rA4 := 3.0584, rA5 := 56.2523, rA6 := 58.7158),
        (rT := 0.8317, rA1 := -120.7638, rA2 := -63.1736, rA3 := 99.5107, rA4 := 6.4400, rA5 := 59.5803, rA6 := 57.3266),
        (rT := 1.1090, rA1 := -121.2340, rA2 := -63.1574, rA3 := 98.6957, rA4 := 10.6204, rA5 := 63.6945, rA6 := 55.6092),
        (rT := 1.3863, rA1 := -121.7582, rA2 := -63.1394, rA3 := 97.7873, rA4 := 15.2801, rA5 := 68.2805, rA6 := 53.6950),
        (rT := 1.6637, rA1 := -122.3003, rA2 := -63.1208, rA3 := 96.8478, rA4 := 20.0996, rA5 := 73.0236, rA6 := 51.7151),
        (rT := 1.9407, rA1 := -122.8245, rA2 := -63.1028, rA3 := 95.9394, rA4 := 24.7593, rA5 := 77.6095, rA6 := 49.8008),
        (rT := 2.2180, rA1 := -123.2947, rA2 := -63.0867, rA3 := 95.1245, rA4 := 28.9397, rA5 := 81.7237, rA6 := 48.0834),
        (rT := 2.4953, rA1 := -123.6751, rA2 := -63.0736, rA3 := 94.4653, rA4 := 32.3213, rA5 := 85.0518, rA6 := 46.6942),
        (rT := 2.7727, rA1 := -123.9297, rA2 := -63.0649, rA3 := 94.0240, rA4 := 34.5845, rA5 := 87.2792, rA6 := 45.7644),
        (rT := 3.0500, rA1 := -124.0225, rA2 := -63.0617, rA3 := 93.8631, rA4 := 35.4100, rA5 := 88.0916, rA6 := 45.4253),
        (rT := 3.1500, rA1 := -124.0227, rA2 := -62.7120, rA3 := 94.1541, rA4 := 35.4756, rA5 := 88.0225, rA6 := 45.3131),
        (rT := 3.2500, rA1 := -124.0229, rA2 := -62.1973, rA3 := 94.5779, rA4 := 35.5837, rA5 := 87.8611, rA6 := 45.0952),
        (rT := 3.3500, rA1 := -124.0230, rA2 := -61.9441, rA3 := 94.7757, rA4 := 35.6709, rA5 := 87.6282, rA6 := 44.8479),
        (rT := 3.4500, rA1 := -124.0229, rA2 := -61.7412, rA3 := 94.9258, rA4 := 35.7491, rA5 := 87.3526, rA6 := 44.5802),
        (rT := 3.5500, rA1 := -124.0229, rA2 := -61.5108, rA3 := 95.0942, rA4 := 35.8058, rA5 := 87.0727, rA6 := 44.3314),
        (rT := 3.6500, rA1 := -124.0229, rA2 := -61.2786, rA3 := 95.2593, rA4 := 35.8504, rA5 := 86.7809, rA6 := 44.0868),
        (rT := 3.7500, rA1 := -124.0229, rA2 := -61.0440, rA3 := 95.4214, rA4 := 35.8877, rA5 := 86.4862, rA6 := 43.8484),
        (rT := 3.8500, rA1 := -124.0229, rA2 := -60.8069, rA3 := 95.5807, rA4 := 35.9201, rA5 := 86.1766, rA6 := 43.6056),
        (rT := 3.9500, rA1 := -124.0229, rA2 := -60.5063, rA3 := 95.7751, rA4 := 35.9594, rA5 := 85.7503, rA6 := 43.2784),
        (rT := 4.0500, rA1 := -124.0229, rA2 := -60.3250, rA3 := 95.8907, rA4 := 35.9822, rA5 := 85.4859, rA6 := 43.0775),
        (* op 7 R1_PARK - traj_robot1_R1_PARK *)
        (rT := 0.0000, rA1 := -124.0229, rA2 := -60.3250, rA3 := 95.8907, rA4 := 35.9822, rA5 := 85.4859, rA6 := 43.0775),
        (rT := 0.2863, rA1 := -125.6247, rA2 := -60.4541, rA3 := 95.8014, rA4 := 35.9822, rA5 := 85.4859, rA6 := 43.0775),
        (rT := 0.5727, rA1 := -129.8294, rA2 := -60.7871, rA3 := 95.5713, rA4 := 35.9822, rA5 := 85.4859, rA6 := 43.0775),
        (rT := 0.8590, rA1 := -135.7360, rA2 := -61.2426, rA3 := 95.2570, rA4 := 35.9822, rA5 := 85.4859, rA6 := 43.0775),
        (rT := 1.1453, rA1 := -142.4435, rA2 := -61.7391, rA3 := 94.9151, rA4 := 35.9822, rA5 := 85.4859, rA6 := 43.0775),
        (rT := 1.4317, rA1 := -149.0509, rA2 := -62.1950, rA3 := 94.6020, rA4 := 35.9822, rA5 := 85.4859, rA6 := 43.0775),
        (rT := 1.7180, rA1 := -154.6572, rA2 := -62.5290, rA3 := 94.3745, rA4 := 35.9822, rA5 := 85.4859, rA6 := 43.0775),
        (rT := 2.0047, rA1 := -158.3613, rA2 := -62.6594, rA3 := 94.2891, rA4 := 35.9822, rA5 := 85.4859, rA6 := 43.0775),
        (rT := 2.0880, rA1 := -160.5075, rA2 := -61.5043, rA3 := 95.1253, rA4 := 35.9822, rA5 := 85.4859, rA6 := 43.0775),
        (rT := 2.1713, rA1 := -158.3613, rA2 := -60.3464, rA3 := 95.9536, rA4 := 35.9822, rA5 := 85.4859, rA6 := 43.0775),
        (* op 8 HOME - traj_robot1_n25 *)
        (rT := 0.0000, rA1 := -158.3613, rA2 := -60.3464, rA3 := 95.9536, rA4 := 35.9822, rA5 := 85.4859, rA6 := 43.0775),
        (rT := 0.2032, rA1 := -158.0833, rA2 := -60.3985, rA3 := 95.9432, rA4 := 35.9190, rA5 := 85.3358, rA6 := 43.0018),
        (rT := 0.4062, rA1 := -157.2676, rA2 := -60.5512, rA3 := 95.9125, rA4 := 35.7336, rA5 := 84.8955, rA6 := 42.7800),
        (rT := 0.6095, rA1 := -155.9418, rA2 := -60.7995, rA3 := 95.8626, rA4 := 35.4324, rA5 := 84.1798, rA6 := 42.4193),
        (rT := 0.8127, rA1 := -154.1335, rA2 := -61.1381, rA3 := 95.7947, rA4 := 35.0215, rA5 := 83.2037, rA6 := 41.9274),
        (rT := 1.0160, rA1 := -151.8703, rA2 := -61.5619, rA3 := 95.7096, rA4 := 34.5073, rA5 := 81.9819, rA6 := 41.3118),
        (rT := 1.2190, rA1 := -149.1796, rA2 := -62.0657, rA3 := 95.6084, rA4 := 33.8959, rA5 := 80.5295, rA6 := 40.5799),
        (rT := 1.4222, rA1 := -146.0892, rA2 := -62.6444, rA3 := 95.4922, rA4 := 33.1937, rA5 := 78.8612, rA6 := 39.7392),
        (rT := 1.6255, rA1 := -142.6265, rA2 := -63.2928, rA3 := 95.3621, rA4 := 32.4070, rA5 := 76.9920, rA6 := 38.7973),
        (rT := 1.8288, rA1 := -138.8192, rA2 := -64.0057, rA3 := 95.2189, rA4 := 31.5419, rA5 := 74.9368, rA6 := 37.7616),
        (rT := 2.0317, rA1 := -134.6948, rA2 := -64.7780, rA3 := 95.0639, rA4 := 30.6048, rA5 := 72.7103, rA6 := 36.6397),
        (rT := 2.2350, rA1 := -130.2809, rA2 := -65.6046, rA3 := 94.8979, rA4 := 29.6018, rA5 := 70.3276, rA6 := 35.4390),
        (rT := 2.4382, rA1 := -125.6050, rA2 := -66.4801, rA3 := 94.7221, rA4 := 28.5394, rA5 := 67.8035, rA6 := 34.1671),
        (rT := 2.6415, rA1 := -120.6948, rA2 := -67.3996, rA3 := 94.5375, rA4 := 27.4237, rA5 := 65.1529, rA6 := 32.8314),
        (rT := 2.8445, rA1 := -115.5777, rA2 := -68.3578, rA3 := 94.3452, rA4 := 26.2611, rA5 := 62.3907, rA6 := 31.4395),
        (rT := 3.0478, rA1 := -110.2815, rA2 := -69.3495, rA3 := 94.1460, rA4 := 25.0577, rA5 := 59.5317, rA6 := 29.9988),
        (rT := 3.2510, rA1 := -104.8336, rA2 := -70.3696, rA3 := 93.9412, rA4 := 23.8198, rA5 := 56.5908, rA6 := 28.5168),
        (rT := 3.4542, rA1 := -99.2616, rA2 := -71.4130, rA3 := 93.7317, rA4 := 22.5538, rA5 := 53.5830, rA6 := 27.0012),
        (rT := 3.6572, rA1 := -93.5931, rA2 := -72.4744, rA3 := 93.5186, rA4 := 21.2658, rA5 := 50.5230, rA6 := 25.4592),
        (rT := 3.8605, rA1 := -87.8557, rA2 := -73.5488, rA3 := 93.3029, rA4 := 19.9622, rA5 := 47.4259, rA6 := 23.8985),
        (rT := 4.0637, rA1 := -82.0769, rA2 := -74.6309, rA3 := 93.0857, rA4 := 18.6492, rA5 := 44.3064, rA6 := 22.3266),
        (rT := 4.2668, rA1 := -76.2844, rA2 := -75.7155, rA3 := 92.8679, rA4 := 17.3330, rA5 := 41.1795, rA6 := 20.7509),
        (rT := 4.4700, rA1 := -70.5056, rA2 := -76.7976, rA3 := 92.6507, rA4 := 16.0200, rA5 := 38.0600, rA6 := 19.1789),
        (rT := 4.6732, rA1 := -64.7682, rA2 := -77.8720, rA3 := 92.4350, rA4 := 14.7163, rA5 := 34.9629, rA6 := 17.6183),
        (rT := 4.8765, rA1 := -59.0997, rA2 := -78.9334, rA3 := 92.2219, rA4 := 13.4284, rA5 := 31.9029, rA6 := 16.0763),
        (rT := 5.0795, rA1 := -53.5277, rA2 := -79.9768, rA3 := 92.0124, rA4 := 12.1623, rA5 := 28.8951, rA6 := 14.5606),
        (rT := 5.2828, rA1 := -48.0798, rA2 := -80.9969, rA3 := 91.8076, rA4 := 10.9245, rA5 := 25.9542, rA6 := 13.0787),
        (rT := 5.4860, rA1 := -42.7836, rA2 := -81.9887, rA3 := 91.6085, rA4 := 9.7211, rA5 := 23.0952, rA6 := 11.6380),
        (rT := 5.6892, rA1 := -37.6666, rA2 := -82.9468, rA3 := 91.4161, rA4 := 8.5584, rA5 := 20.3330, rA6 := 10.2461),
        (rT := 5.8922, rA1 := -32.7563, rA2 := -83.8663, rA3 := 91.2315, rA4 := 7.4427, rA5 := 17.6824, rA6 := 8.9104),
        (rT := 6.0955, rA1 := -28.0805, rA2 := -84.7419, rA3 := 91.0557, rA4 := 6.3803, rA5 := 15.1583, rA6 := 7.6385),
        (rT := 6.2987, rA1 := -23.6665, rA2 := -85.5684, rA3 := 90.8897, rA4 := 5.3774, rA5 := 12.7756, rA6 := 6.4378),
        (rT := 6.5020, rA1 := -19.5421, rA2 := -86.3407, rA3 := 90.7347, rA4 := 4.4403, rA5 := 10.5491, rA6 := 5.3159),
        (rT := 6.7050, rA1 := -15.7348, rA2 := -87.0536, rA3 := 90.5916, rA4 := 3.5752, rA5 := 8.4939, rA6 := 4.2802),
        (rT := 6.9082, rA1 := -12.2721, rA2 := -87.7020, rA3 := 90.4614, rA4 := 2.7884, rA5 := 6.6247, rA6 := 3.3383),
        (rT := 7.1115, rA1 := -9.1817, rA2 := -88.2807, rA3 := 90.3452, rA4 := 2.0862, rA5 := 4.9564, rA6 := 2.4976),
        (rT := 7.3147, rA1 := -6.4911, rA2 := -88.7845, rA3 := 90.2440, rA4 := 1.4749, rA5 := 3.5040, rA6 := 1.7657),
        (rT := 7.5177, rA1 := -4.2278, rA2 := -89.2083, rA3 := 90.1589, rA4 := 0.9606, rA5 := 2.2822, rA6 := 1.1500),
        (rT := 7.7210, rA1 := -2.4195, rA2 := -89.5469, rA3 := 90.0910, rA4 := 0.5497, rA5 := 1.3061, rA6 := 0.6582),
        (rT := 7.9242, rA1 := -1.0937, rA2 := -89.7952, rA3 := 90.0411, rA4 := 0.2485, rA5 := 0.5904, rA6 := 0.2975),
        (rT := 8.1273, rA1 := -0.2780, rA2 := -89.9479, rA3 := 90.0105, rA4 := 0.0632, rA5 := 0.1501, rA6 := 0.0756),
        (rT := 8.3305, rA1 := 0.0000, rA2 := -90.0000, rA3 := 90.0000, rA4 := 0.0000, rA5 := 0.0000, rA6 := 0.0000)
    ];
END_VAR
END_NAMESPACE

(* ---- FB_JointAngleEncoder.st ---- *)
(*
 * FB_JointAngleEncoder
 * Device simulator R1 (robot1), cell welding_cell_2_small. Generated by bt2plc 0.1.0.
 *
 * Encodes six KUKA robot joint angles (REAL degrees) into the VASS Option area
 * as scaled fixed-point INTs (0.02 deg per count, big-endian byte order).
 *
 * Encoding per encoding.md:
 *   count = ROUND(angle_deg / 0.02)   clamped to [-32768, +32767]
 *   Byte layout: big-endian (high byte first) in each 2-byte pair
 *
 * Output abyOption = Option area aVassInputData[16..27], 2 bytes per axis
 * (PLC_PRG copies it into the robot -> PLC telegram):
 *   abyOption[0-1]  = bytes 16-17 = A1,  abyOption[2-3]   = bytes 18-19 = A2,
 *   abyOption[4-5]  = bytes 20-21 = A3,  abyOption[6-7]   = bytes 22-23 = A4,
 *   abyOption[8-9]  = bytes 24-25 = A5,  abyOption[10-11] = bytes 26-27 = A6
 *)

FUNCTION_BLOCK FB_JointAngleEncoder
VAR_INPUT
    rA1_deg     : REAL := 0.0;      (* Axis 1 angle in degrees *)
    rA2_deg     : REAL := 0.0;      (* Axis 2 angle in degrees *)
    rA3_deg     : REAL := 0.0;      (* Axis 3 angle in degrees *)
    rA4_deg     : REAL := 0.0;      (* Axis 4 angle in degrees *)
    rA5_deg     : REAL := 0.0;      (* Axis 5 angle in degrees *)
    rA6_deg     : REAL := 0.0;      (* Axis 6 angle in degrees *)
END_VAR

VAR_OUTPUT
    (* Encoded INT values (for monitoring/debug) *)
    iA1_count   : INT;
    iA2_count   : INT;
    iA3_count   : INT;
    iA4_count   : INT;
    iA5_count   : INT;
    iA6_count   : INT;

    (* Option area bytes 16..27 of the robot -> PLC telegram, big-endian A1..A6 *)
    abyOption   : ARRAY[0..11] OF BYTE;
END_VAR

VAR CONSTANT
    SCALE_FACTOR    : REAL := 0.02;     (* degrees per count *)
    INV_SCALE       : REAL := 50.0;     (* 1/0.02 = 50, multiply for speed *)
    COUNT_MAX       : DINT := 32767;
    COUNT_MIN       : DINT := -32768;
END_VAR

VAR
    _arDeg      : ARRAY[1..6] OF REAL;
    _aiCount    : ARRAY[1..6] OF INT;
    _diTemp     : DINT;
    _wTemp      : WORD;
    _i          : INT;
END_VAR
(*
 * FB_JointAngleEncoder - Implementation
 *
 * Converts 6x REAL degree angles to scaled INT counts (0.02 deg per count)
 * and writes them big-endian into abyOption[0..11] (telegram bytes 16..27).
 *
 * Conversion:  count = ROUND(angle / 0.02)  clamped to INT range
 * Byte order:  Big-endian (high byte at lower address) per S7/PROFINET convention
 * Two's complement is formed in DINT (count + 65536 for negative counts), so no
 * bit operation is applied to a signed type.
 *)

_arDeg[1] := rA1_deg;
_arDeg[2] := rA2_deg;
_arDeg[3] := rA3_deg;
_arDeg[4] := rA4_deg;
_arDeg[5] := rA5_deg;
_arDeg[6] := rA6_deg;

FOR _i := 1 TO 6 DO
    (* === Scale and clamp === *)
    _diTemp := REAL_TO_DINT(LIMIT(REAL#-32768.0, _arDeg[_i] * INV_SCALE, REAL#32767.0));
    IF _diTemp > COUNT_MAX THEN _diTemp := COUNT_MAX; END_IF
    IF _diTemp < COUNT_MIN THEN _diTemp := COUNT_MIN; END_IF
    _aiCount[_i] := DINT_TO_INT(_diTemp);

    (* === Big-endian into the Option area: high byte first === *)
    IF _diTemp < 0 THEN
        _diTemp := _diTemp + 65536;
    END_IF
    _wTemp := DINT_TO_WORD(_diTemp);
    abyOption[2 * (_i - 1)] := WORD_TO_BYTE(SHR(_wTemp, 8));
    abyOption[2 * (_i - 1) + 1] := WORD_TO_BYTE(_wTemp AND WORD#16#FF);
END_FOR

iA1_count := _aiCount[1];
iA2_count := _aiCount[2];
iA3_count := _aiCount[3];
iA4_count := _aiCount[4];
iA5_count := _aiCount[5];
iA6_count := _aiCount[6];
END_FUNCTION_BLOCK

(* ---- FB_PROFIsafe_Simulator.st ---- *)
(*
 * FB_PROFIsafe_Simulator
 * Device simulator R1 (robot1), cell welding_cell_2_small. Generated by bt2plc 0.1.0.
 *
 * Simulates the PROFIsafe protocol layer for the FDIO64 module (Slot 1).
 * In a real KUKA controller, the PROFIsafe stack handles CRC generation,
 * sequence counters, and watchdog monitoring.
 *
 * For simulation purposes, this FB:
 * - Monitors the safe output bytes from the PLC (abySafeOut = copy of GVL_IO.bySafeOut0..7)
 * - Provides a "communication OK" flag
 *
 * IMPORTANT: This does NOT provide real functional safety!
 * It only generates data patterns that allow the PLC's PROFIsafe stack
 * to accept the device as communicating. For real safety testing,
 * you need a certified PROFIsafe device or test equipment.
 *
 * PROFIsafe frame structure per IEC 61784-3-3:
 *   [User Data (8 bytes)] [Status/Control (1 byte)] [CRC (3 bytes)]
 *
 * Status byte bits (F_Input from device):
 *   Bit 0: Toggle bit (alternates each cycle)
 *   Bit 1: Reserved
 *   Bit 2: Data valid
 *   Bit 3-7: Reserved / Sequence counter
 *
 * Control byte bits (F_Output from controller):
 *   Bit 0: Toggle bit
 *   Bit 1: Activate device
 *   Bit 2: Reserved
 *   Bit 3-7: Reserved
 *)

FUNCTION_BLOCK FB_PROFIsafe_Simulator
VAR_INPUT
    bEnable         : BOOL := TRUE;
    dwF_Source_Add  : DWORD := DWORD#1;     (* F_Source_Add from parameterization *)
    dwF_Dest_Add    : DWORD := DWORD#1;     (* F_Dest_Add from parameterization *)
    tF_WD_Time      : TIME := T#500MS;      (* Watchdog time *)
    abySafeOut      : ARRAY[0..7] OF BYTE;  (* Safe outputs PLC -> robot (GVL_IO.bySafeOut0..7) *)
END_VAR

VAR_OUTPUT
    bCommOK         : BOOL;                 (* PROFIsafe communication established *)
    bDataValid      : BOOL;                 (* Safe data is valid *)
    bWatchdogError  : BOOL;                 (* Watchdog timeout *)
END_VAR

VAR
    _bToggleBit     : BOOL;                 (* Toggle bit for sequence *)
    _nSeqCounter    : BYTE;                 (* Sequence counter 0-31 *)
    _nCycleCount    : UDINT;                (* Absolute cycle counter *)

    (* Watchdog *)
    _tonWatchdog    : TON;
    _bPLCSafeActive : BOOL;

    (* CRC calculation helper *)
    _dwCrcSeed      : DWORD;
END_VAR
(*
 * FB_PROFIsafe_Simulator - Implementation
 * Works on the input image abySafeOut (PLC_PRG copies GVL_IO.bySafeOut0..7).
 *)

IF NOT bEnable THEN
    bCommOK := FALSE;
    bDataValid := FALSE;
    RETURN;
END_IF

IF _nCycleCount < UDINT#4000000000 THEN
    _nCycleCount := _nCycleCount + 1;
ELSE
    _nCycleCount := 0;
END_IF

(* ============================================================================
   MONITOR PLC SAFE OUTPUT DATA
   ============================================================================ *)
_bPLCSafeActive := (abySafeOut[0] <> BYTE#0) OR (abySafeOut[1] <> BYTE#0);

(* Watchdog *)
_tonWatchdog(IN := NOT _bPLCSafeActive, PT := tF_WD_Time);
bWatchdogError := _tonWatchdog.Q;

bCommOK := _bPLCSafeActive AND NOT bWatchdogError;
bDataValid := bCommOK;
END_FUNCTION_BLOCK

(* ---- FB_ProgramPlayer.st ---- *)
(*
 * FB_ProgramPlayer
 * Device simulator R1 (robot1), cell welding_cell_2_small, tree bt_1790934549_welding_cell_2_small. Generated by bt2plc 0.1.0.
 *
 * Plays the bt2plc robot program (GVL_Program) for PROD_FOLGE, or a blind joint
 * move to the home pose for HOME_FOLGE. Robot side of the zone protocol, per op k
 * with mask M = GVL_Program.aOps[k].dwZoneMask:
 *   1  wStep := k                          (also for M = 0)
 *   2  if M <> 0: REQUEST := M             (same call / telegram as wStep)
 *   3  if M <> 0: wait (GRANT AND M) = M
 *   4  start delay; trajectory (x rVelScale x override); hold
 *   5  if M <> 0: REQUEST := 0
 *   6  if M <> 0: wait (GRANT AND M) = 0   (4-phase, before the next REQUEST)
 *   7  next op; after the last op: bDone, wStep := 0 (same call)
 *
 * Timing: all times are REAL seconds accumulated from rDt (seconds per call, the
 * device task interval). Motion time advances by rDt * rRate * rVelScale, delay and
 * hold by rDt (the override does not scale dwell times). No TIME() / TON is used.
 * Zero-time transitions fall through within one call (at most N_MAX_TRANSITIONS),
 * but wStep changes at most once per call, so every step is visible to the head PLC.
 * Joints (deg) are linearly interpolated between waypoints and published as rA1..rA6_deg.
 * Abort (bAbort level while busy): REQUEST := 0, wStep := 0, the pose is held.
 * The robot powers up at GVL_Program.arHomeDeg.
 *)

FUNCTION_BLOCK FB_ProgramPlayer
VAR_INPUT
    bStart          : BOOL;                 (* Rising edge: start wJob *)
    wJob            : WORD;                 (* Folge to play: PROD_FOLGE or HOME_FOLGE *)
    bAbort          : BOOL;                 (* Level: stop / cancel / drives off / E-stop *)
    dwGrant         : DWORD;                (* Zone GRANT bits from the head PLC *)
    rRate           : REAL := 1.0;          (* Speed override factor (1.0 = 100 %) *)
    rDt             : REAL := 0.02;         (* Seconds per call (task interval) *)
END_VAR

VAR_OUTPUT
    eState          : E_PlayerState;        (* Current state *)
    bBusy           : BOOL;                 (* Program running *)
    bDone           : BOOL;                 (* Latched until next start *)
    bError          : BOOL;                 (* Latched until next start *)
    wErrorCode      : WORD;                 (* Error code, GVL_Program.ERR_xxx *)
    wWarningCode    : WORD;                 (* Warning code, GVL_Program.WARN_xxx, latched until next start *)
    wStep           : WORD;                 (* 1-based op index, 0 = none *)
    dwRequest       : DWORD;                (* Zone REQUEST bits to the head PLC *)
    bAtHome         : BOOL;                 (* All joints within R_AT_HOME_TOL_DEG of arHomeDeg *)
    rA1_deg         : REAL;                 (* Axis 1 angle *)
    rA2_deg         : REAL;                 (* Axis 2 angle *)
    rA3_deg         : REAL;                 (* Axis 3 angle *)
    rA4_deg         : REAL;                 (* Axis 4 angle *)
    rA5_deg         : REAL;                 (* Axis 5 angle *)
    rA6_deg         : REAL;                 (* Axis 6 angle *)
END_VAR

VAR CONSTANT
    N_MAX_TRANSITIONS : INT := 8;           (* Fall-through bound per call *)
END_VAR

VAR
    _eState         : E_PlayerState := E_PlayerState#PS_IDLE;
    _rtrigStart     : R_TRIG;
    _bFirstCall     : BOOL := TRUE;

    (* === Current op === *)
    _nOp            : INT;                  (* 1-based op index, 0 = HOME_FOLGE move *)
    _dwMask         : DWORD;                (* Zone mask of the current op *)
    _bHomeMove      : BOOL;                 (* Current move is a blind home move *)
    _nWp            : INT;                  (* Current waypoint segment start *)
    _nLast          : INT;                  (* Last waypoint of the current op, 0 = none *)
    _rVel           : REAL;                 (* Velocity scale of the current move *)

    (* === Time (s) === *)
    _rDtCall        : REAL;                 (* rDt limited to 0..1 s *)
    _rRateCall      : REAL;                 (* rRate limited to >= 0 *)
    _rT             : REAL;                 (* Motion time since move start *)
    _rTimer         : REAL;                 (* Delay / hold timer *)
    _rDur           : REAL;                 (* Duration of the blind home move *)
    _rAlpha         : REAL;                 (* Interpolation factor 0..1 *)
    _rSpan          : REAL;                 (* Waypoint segment duration *)

    (* === Pose (deg) === *)
    _arQ            : ARRAY[1..6] OF REAL;  (* Current joint angles *)
    _arQ0           : ARRAY[1..6] OF REAL;  (* Pose at the start of a blind home move *)
    _arQa           : ARRAY[1..6] OF REAL;  (* Segment start waypoint *)
    _arQb           : ARRAY[1..6] OF REAL;  (* Segment end waypoint *)

    (* === Fall-through === *)
    _nPass          : INT;
    _bAdvance       : BOOL;                 (* A transition happened in this pass *)
    _bStepSet       : BOOL;                 (* wStep changed in this call *)
    _bMoveDone      : BOOL;
    _i              : INT;
END_VAR
(*
 * FB_ProgramPlayer - Implementation
 *)

(* ============================================================================
   INIT - the robot powers up at the home pose
   ============================================================================ *)
IF _bFirstCall THEN
    FOR _i := 1 TO 6 DO
        _arQ[_i] := GVL_Program.arHomeDeg[_i];
    END_FOR
    _bFirstCall := FALSE;
END_IF

_rDtCall := LIMIT(0.0, rDt, 1.0);
_rRateCall := MAX(rRate, 0.0);
_rtrigStart(CLK := bStart);

(* ============================================================================
   ABORT - stop / cancel / drives off / E-stop: REQUEST := 0, wStep := 0, hold pose
   ============================================================================ *)
IF bAbort AND bBusy THEN
    _eState := E_PlayerState#PS_IDLE;
    bBusy := FALSE;
    wStep := WORD#0;
    dwRequest := DWORD#0;
END_IF

(* ============================================================================
   CLOCK - advance the timer of the state that is active at the start of the call
   (a state entered during this call starts counting with the next call)
   ============================================================================ *)
IF _eState = E_PlayerState#PS_DELAY OR _eState = E_PlayerState#PS_HOLD THEN
    _rTimer := _rTimer + _rDtCall;
ELSIF _eState = E_PlayerState#PS_MOVE THEN
    _rT := _rT + _rDtCall * _rRateCall * _rVel;
END_IF

(* ============================================================================
   START
   ============================================================================ *)
IF _rtrigStart.Q AND NOT bBusy AND NOT bAbort THEN
    bDone := FALSE;
    bError := FALSE;
    wErrorCode := WORD#0;
    wWarningCode := WORD#0;
    wStep := WORD#0;
    dwRequest := DWORD#0;
    _nOp := 0;
    _dwMask := DWORD#0;
    _rT := 0.0;
    _rTimer := 0.0;
    IF wJob = GVL_Program.HOME_FOLGE THEN
        (* Blind joint move from the current pose to arHomeDeg: no step, no zones *)
        FOR _i := 1 TO 6 DO
            _arQ0[_i] := _arQ[_i];
        END_FOR
        _bHomeMove := TRUE;
        _nLast := 0;
        _rVel := 1.0;
        _rDur := GVL_Program.R_HOME_S;
        bBusy := TRUE;
        _eState := E_PlayerState#PS_MOVE;
    ELSIF wJob = GVL_Program.PROD_FOLGE AND GVL_Program.N_OPS > 0 THEN
        bBusy := TRUE;
        _eState := E_PlayerState#PS_NEXT_OP;
    ELSE
        wErrorCode := GVL_Program.ERR_UNKNOWN_FOLGE;
        _eState := E_PlayerState#PS_ERROR;
    END_IF
END_IF

(* ============================================================================
   STATE MACHINE - falls through zero-time transitions (bounded)
   ============================================================================ *)
_bStepSet := FALSE;
FOR _nPass := 1 TO N_MAX_TRANSITIONS DO
    _bAdvance := FALSE;

    CASE _eState OF

    E_PlayerState#PS_IDLE:
        bBusy := FALSE;
        wStep := WORD#0;
        dwRequest := DWORD#0;

    E_PlayerState#PS_NEXT_OP:
        (* wStep changes at most once per call: the head checks step + 1 per telegram *)
        IF NOT _bStepSet THEN
            _nOp := _nOp + 1;
            IF _nOp > GVL_Program.N_OPS THEN
                _eState := E_PlayerState#PS_DONE;
            ELSE
                wStep := INT_TO_WORD(_nOp);
                _bStepSet := TRUE;
                _dwMask := GVL_Program.aOps[_nOp].dwZoneMask;
                IF _dwMask <> DWORD#0 THEN
                    dwRequest := _dwMask;           (* same telegram as wStep *)
                    _eState := E_PlayerState#PS_WAIT_GRANT;
                ELSE
                    _rTimer := 0.0;
                    _eState := E_PlayerState#PS_DELAY;
                END_IF
            END_IF
            _bAdvance := TRUE;
        END_IF

    E_PlayerState#PS_WAIT_GRANT:
        IF (dwGrant AND _dwMask) = _dwMask THEN
            _rTimer := 0.0;
            _eState := E_PlayerState#PS_DELAY;
            _bAdvance := TRUE;
        END_IF

    E_PlayerState#PS_DELAY:
        IF _rTimer >= GVL_Program.aOps[_nOp].rDelay_s THEN
            (* Begin the motion of op _nOp *)
            _rT := 0.0;
            _rVel := GVL_Program.aOps[_nOp].rVelScale;
            IF _rVel <= 0.0 THEN
                _rVel := 1.0;
            END_IF
            _bHomeMove := GVL_Program.aOps[_nOp].bBlindHome;
            IF _bHomeMove THEN
                FOR _i := 1 TO 6 DO
                    _arQ0[_i] := _arQ[_i];
                END_FOR
                _rDur := GVL_Program.R_HOME_S;
                _nLast := 0;
            ELSE
                _nWp := GVL_Program.aOps[_nOp].nFirstWp;
                _nLast := GVL_Program.aOps[_nOp].nLastWp;
                IF _nWp < 1 OR _nLast < _nWp OR _nLast > GVL_Program.N_WP THEN
                    _nLast := 0;                    (* no valid trajectory: zero-length move *)
                ELSE
                    (* Start deviation: the trajectory should start at the current pose *)
                    _arQa[1] := GVL_Program.aWp[_nWp].rA1;
                    _arQa[2] := GVL_Program.aWp[_nWp].rA2;
                    _arQa[3] := GVL_Program.aWp[_nWp].rA3;
                    _arQa[4] := GVL_Program.aWp[_nWp].rA4;
                    _arQa[5] := GVL_Program.aWp[_nWp].rA5;
                    _arQa[6] := GVL_Program.aWp[_nWp].rA6;
                    FOR _i := 1 TO 6 DO
                        IF ABS(_arQ[_i] - _arQa[_i]) > GVL_Program.R_START_TOL_DEG THEN
                            wWarningCode := GVL_Program.WARN_START_DEVIATION;
                        END_IF
                    END_FOR
                END_IF
            END_IF
            _eState := E_PlayerState#PS_MOVE;
            _bAdvance := TRUE;
        END_IF

    E_PlayerState#PS_MOVE:
        _bMoveDone := FALSE;
        IF _bHomeMove THEN
            (* Blind joint move: linear in joint space over R_HOME_S *)
            IF _rDur > 0.0 THEN
                _rAlpha := LIMIT(0.0, _rT / _rDur, 1.0);
            ELSE
                _rAlpha := 1.0;
            END_IF
            FOR _i := 1 TO 6 DO
                _arQ[_i] := _arQ0[_i] + _rAlpha * (GVL_Program.arHomeDeg[_i] - _arQ0[_i]);
            END_FOR
            _bMoveDone := _rAlpha >= 1.0;
        ELSIF _nLast < 1 THEN
            _bMoveDone := TRUE;
        ELSE
            (* Trajectory: find the segment [_nWp, _nWp + 1] that contains _rT *)
            WHILE _nWp < _nLast DO
                IF GVL_Program.aWp[_nWp + 1].rT <= _rT THEN
                    _nWp := _nWp + 1;
                ELSE
                    EXIT;
                END_IF
            END_WHILE
            _arQa[1] := GVL_Program.aWp[_nWp].rA1;
            _arQa[2] := GVL_Program.aWp[_nWp].rA2;
            _arQa[3] := GVL_Program.aWp[_nWp].rA3;
            _arQa[4] := GVL_Program.aWp[_nWp].rA4;
            _arQa[5] := GVL_Program.aWp[_nWp].rA5;
            _arQa[6] := GVL_Program.aWp[_nWp].rA6;
            IF _nWp >= _nLast THEN
                FOR _i := 1 TO 6 DO
                    _arQ[_i] := _arQa[_i];
                END_FOR
                _bMoveDone := TRUE;
            ELSE
                _arQb[1] := GVL_Program.aWp[_nWp + 1].rA1;
                _arQb[2] := GVL_Program.aWp[_nWp + 1].rA2;
                _arQb[3] := GVL_Program.aWp[_nWp + 1].rA3;
                _arQb[4] := GVL_Program.aWp[_nWp + 1].rA4;
                _arQb[5] := GVL_Program.aWp[_nWp + 1].rA5;
                _arQb[6] := GVL_Program.aWp[_nWp + 1].rA6;
                _rSpan := GVL_Program.aWp[_nWp + 1].rT - GVL_Program.aWp[_nWp].rT;
                IF _rSpan > 0.0 THEN
                    _rAlpha := LIMIT(0.0, (_rT - GVL_Program.aWp[_nWp].rT) / _rSpan, 1.0);
                ELSE
                    _rAlpha := 1.0;
                END_IF
                FOR _i := 1 TO 6 DO
                    _arQ[_i] := _arQa[_i] + _rAlpha * (_arQb[_i] - _arQa[_i]);
                END_FOR
            END_IF
        END_IF
        IF _bMoveDone THEN
            IF _nOp = 0 THEN
                _eState := E_PlayerState#PS_DONE;   (* HOME_FOLGE finished *)
            ELSE
                _rTimer := 0.0;
                _eState := E_PlayerState#PS_HOLD;
            END_IF
            _bAdvance := TRUE;
        END_IF

    E_PlayerState#PS_HOLD:
        IF _rTimer >= GVL_Program.aOps[_nOp].rHold_s THEN
            IF _dwMask <> DWORD#0 THEN
                dwRequest := DWORD#0;
                _eState := E_PlayerState#PS_WAIT_RELEASE;
            ELSE
                _eState := E_PlayerState#PS_NEXT_OP;
            END_IF
            _bAdvance := TRUE;
        END_IF

    E_PlayerState#PS_WAIT_RELEASE:
        (* 4-phase: the GRANT must drop before the next REQUEST *)
        IF (dwGrant AND _dwMask) = DWORD#0 THEN
            _eState := E_PlayerState#PS_NEXT_OP;
            _bAdvance := TRUE;
        END_IF

    E_PlayerState#PS_DONE:
        bBusy := FALSE;
        bDone := TRUE;
        wStep := WORD#0;
        dwRequest := DWORD#0;
        _eState := E_PlayerState#PS_IDLE;

    E_PlayerState#PS_ERROR:
        bBusy := FALSE;
        bError := TRUE;
        wStep := WORD#0;
        dwRequest := DWORD#0;
        _eState := E_PlayerState#PS_IDLE;

    END_CASE

    IF NOT _bAdvance THEN
        EXIT;
    END_IF
END_FOR

(* ============================================================================
   PUBLISH
   ============================================================================ *)
bAtHome := TRUE;
FOR _i := 1 TO 6 DO
    IF ABS(_arQ[_i] - GVL_Program.arHomeDeg[_i]) > GVL_Program.R_AT_HOME_TOL_DEG THEN
        bAtHome := FALSE;
    END_IF
END_FOR
rA1_deg := _arQ[1];
rA2_deg := _arQ[2];
rA3_deg := _arQ[3];
rA4_deg := _arQ[4];
rA5_deg := _arQ[5];
rA6_deg := _arQ[6];
eState := _eState;
END_FUNCTION_BLOCK

(* ---- FB_VASS_DeviceSimulator.st ---- *)
(*
 * FB_VASS_DeviceSimulator
 * Device simulator R1 (robot1, station kuka-robi1), cell welding_cell_2_small, tree bt_1790934549_welding_cell_2_small.
 * Generated by bt2plc 0.1.0.
 *
 * Simulates a KUKA KR C4 robot responding to VW VASS commands via PROFINET.
 *
 * This FB reads the PLC commands from its input images (PLC -> robot):
 *   aVassOutputData = copy of GVL_IO.aVassOutputData, abySafeOut = GVL_IO.bySafeOut0..7
 * and produces the robot status images (robot -> PLC):
 *   aVassInputData (bytes 16-27 = 0, the joint encoder fills them in PLC_PRG), abySafeIn.
 * PLC_PRG copies the images from / to GVL_IO; this FB never accesses GVL_IO.
 *
 * Job handshake (as the original simulator): drives on after 2 s, EXT mode, Ready,
 * JobRequest edge -> JobAck + job echo (clears ProgFinished), ProgStart edge -> start,
 * Stop/Cancel level -> stop, Reset held 500 ms -> clear error, gripper, speed override.
 * Job execution is delegated to FB_ProgramPlayer (GVL_Program):
 *   PROD_FOLGE: the bt2plc program; PLAN_ID (bytes PLAN_ID_BYTE..+1, latched at job accept)
 *               must equal GVL_Program.PLAN_ID at ProgStart, else ERR_PLAN_MISMATCH, no start.
 *   HOME_FOLGE: blind joint move to arHomeDeg (also on a HomeRequest [0].6 edge while Ready).
 *   other:      ERR_UNKNOWN_FOLGE, no start.
 * Zone protocol: wCurrentStep at bytes STEP_BYTE..+1, REQUEST DWORD LE at REQ_BYTE..+3,
 * GRANT DWORD LE read from bytes GRANT_BYTE..+3 (GVL_Program offsets).
 * At the end ProgRunning := FALSE, ProgFinished := TRUE and step := 0 in the same scan.
 *)

FUNCTION_BLOCK FB_VASS_DeviceSimulator
VAR_INPUT
    bEnable             : BOOL := TRUE;             (* Enable simulation *)
    wRobotID            : WORD := WORD#1;           (* Robot identification number 1-8 *)
    aVassOutputData     : ARRAY[0..31] OF BYTE;     (* VASS telegram PLC -> robot (GVL_IO.aVassOutputData) *)
    abySafeOut          : ARRAY[0..7] OF BYTE;      (* Safe outputs PLC -> robot (GVL_IO.bySafeOut0..7) *)
    rDt                 : REAL := 0.02;             (* Task interval in s (GVL_Program.R_TASK_S) *)
END_VAR

VAR_OUTPUT
    bActive             : BOOL;                     (* Simulator is active *)
    eCurrentMode        : E_RobotMode;              (* Current operating mode *)
    eProgramState       : E_ProgramState;           (* Current program state *)
    bSafetyOK           : BOOL;                     (* Safety system healthy *)
    aVassInputData      : ARRAY[0..31] OF BYTE;     (* VASS telegram robot -> PLC (bytes 16-27 = 0) *)
    abySafeIn           : ARRAY[0..7] OF BYTE;      (* Safe inputs robot -> PLC (GVL_IO.bySafeIn0..7) *)

    (* Joint angles from the program player (deg) *)
    rA1_deg             : REAL;
    rA2_deg             : REAL;
    rA3_deg             : REAL;
    rA4_deg             : REAL;
    rA5_deg             : REAL;
    rA6_deg             : REAL;

    (* Diagnostics *)
    wActiveJob          : WORD;                     (* Accepted job number (Folge) *)
    wCurrentStep        : WORD;                     (* Current op index, 0 = none *)
    wErrorCode          : WORD;                     (* Active error code *)
    dwRequest           : DWORD;                    (* Zone REQUEST bits sent to the head PLC *)
    dwGrant             : DWORD;                    (* Zone GRANT bits received from the head PLC *)
    ePlayerState        : E_PlayerState;            (* State of the program player *)
END_VAR

VAR
    (* === Internal Robot State === *)
    _bDrivesPowered     : BOOL;
    _bInExtMode         : BOOL;
    _bReady             : BOOL;
    _bError             : BOOL;
    _bProgRunning       : BOOL;
    _bAtHome            : BOOL := TRUE;
    _bInPosition        : BOOL := TRUE;
    _bProgFinished      : BOOL;
    _bJobAcknowledged   : BOOL;
    _bGripperClosed     : BOOL;
    _bPartPresent       : BOOL;
    _bPeriphReady       : BOOL := TRUE;

    _wActiveJob         : WORD;
    _wCurrentStep       : WORD;
    _wSpeed             : WORD := WORD#100;
    _wToolNr            : WORD := WORD#1;
    _wErrorCode         : WORD;
    _wWarningCode       : WORD;

    (* Simulated position (0.1mm units) *)
    _iPositionX         : INT := 5000;              (* 500.0 mm *)
    _iPositionY         : INT := 0;
    _iPositionZ         : INT := 10000;             (* 1000.0 mm *)

    (* === Safety State === *)
    _bSafe_DrivesOK     : BOOL := TRUE;
    _bSafe_Stopped      : BOOL := TRUE;
    _bSafe_EStopOK      : BOOL := TRUE;
    _bSafe_GatesClosed  : BOOL := TRUE;
    _bSafe_Fault        : BOOL;
    _bSafe_STO          : BOOL;
    _bSafe_SS1          : BOOL;

    (* PROFIsafe CRC simulation *)
    _bySafeTrailerStatus : BYTE;
    _nSafeCycleCount     : UDINT;

    (* === Timers === *)
    _tonDriveStartup    : TON;                      (* Simulate drive power-on delay *)
    _tonErrorReset      : TON;                      (* Simulate error reset delay *)
    _tonGripperAction   : TON;                      (* Simulate gripper open/close time *)

    (* === Edge Detection === *)
    _rtrigProgStart     : R_TRIG;
    _rtrigProgStop      : R_TRIG;
    _rtrigReset         : R_TRIG;
    _rtrigJobReq        : R_TRIG;
    _rtrigDrivesOn      : R_TRIG;
    _rtrigHome          : R_TRIG;
    _rtrigGripOpen      : R_TRIG;
    _rtrigGripClose     : R_TRIG;
    _rtrigSafeStop1     : R_TRIG;
    _rtrigSafeEStop     : R_TRIG;

    (* === Program player (bt2plc program / blind home) === *)
    _fbPlayer           : FB_ProgramPlayer;
    _bPlayerStart       : BOOL;                     (* Start pulse for the player *)
    _wPlayerJob         : WORD;                     (* Folge passed to the player *)
    _bStartOk           : BOOL;
    _wPlanId            : WORD;                     (* PLAN_ID latched at job accept *)
    _dwGrant            : DWORD;
    _dwRequest          : DWORD;
    _rRate              : REAL;                     (* Speed override factor *)
    _wPlayerWarning     : WORD;                     (* Last player warning (copy on change) *)

    (* === Decoded PLC commands (aVassOutputData bytes 0-1, abySafeOut byte 0) === *)
    _bCmdDrivesOn       : BOOL;                     (* [0].0 Drives on *)
    _bCmdProgStart      : BOOL;                     (* [0].1 Program start *)
    _bCmdProgStop       : BOOL;                     (* [0].2 Program stop *)
    _bCmdProgCancel     : BOOL;                     (* [0].3 Program cancel *)
    _bCmdModeExt        : BOOL;                     (* [0].4 EXT mode request *)
    _bCmdReset          : BOOL;                     (* [0].5 Reset *)
    _bCmdHome           : BOOL;                     (* [0].6 Home request *)
    _bCmdJobReq         : BOOL;                     (* [1].0 Job request *)
    _bCmdGripOpen       : BOOL;                     (* [1].1 Gripper open *)
    _bCmdGripClose      : BOOL;                     (* [1].2 Gripper close *)
    _bCmdSpeedOverride  : BOOL;                     (* [1].4 Apply speed override *)
    _bSafeCmdDriveEnable : BOOL;                    (* Safe [0].0 Drive enable *)
    _bSafeCmdEStop      : BOOL;                     (* Safe [0].1 External E-Stop *)
    _bSafeCmdSS1        : BOOL;                     (* Safe [0].2 Safe Stop 1 *)

    (* === Local working variables === *)
    _wRequestedJob      : WORD;
    _wSpeedCmd          : WORD;
    _nIdx               : INT;
    _i                  : INT;
END_VAR
(*
 * FB_VASS_DeviceSimulator - Implementation
 *
 * Reads commands from aVassOutputData (PLC -> Robot, 32 bytes) and abySafeOut (8 bytes).
 * Writes status to aVassInputData (Robot -> PLC, 32 bytes) and abySafeIn (8 bytes).
 *)

IF NOT bEnable THEN
    bActive := FALSE;
    RETURN;
END_IF

bActive := TRUE;

(* ============================================================================
   SECTION 1: READ PLC COMMANDS from aVassOutputData[0..31]
   Byte 0-1 = Control word, Byte 2-3 = Job number, PLAN_ID / GRANT per GVL_Program
   ============================================================================ *)

(* Decode the control bits into BOOLs (a bare bit access is never passed as a call argument) *)
_bCmdDrivesOn       := aVassOutputData[0].0;
_bCmdProgStart      := aVassOutputData[0].1;
_bCmdProgStop       := aVassOutputData[0].2;
_bCmdProgCancel     := aVassOutputData[0].3;
_bCmdModeExt        := aVassOutputData[0].4;
_bCmdReset          := aVassOutputData[0].5;
_bCmdHome           := aVassOutputData[0].6;
_bCmdJobReq         := aVassOutputData[1].0;
_bCmdGripOpen       := aVassOutputData[1].1;
_bCmdGripClose      := aVassOutputData[1].2;
_bCmdSpeedOverride  := aVassOutputData[1].4;
_bSafeCmdDriveEnable := abySafeOut[0].0;
_bSafeCmdEStop      := abySafeOut[0].1;
_bSafeCmdSS1        := abySafeOut[0].2;

(* Edge detection on control signals - output byte 0 *)
_rtrigDrivesOn(CLK  := _bCmdDrivesOn);
_rtrigProgStart(CLK := _bCmdProgStart);
_rtrigProgStop(CLK  := _bCmdProgStop);
_rtrigReset(CLK     := _bCmdReset);
_rtrigHome(CLK      := _bCmdHome);

(* Output byte 1 *)
_rtrigJobReq(CLK    := _bCmdJobReq);
_rtrigGripOpen(CLK  := _bCmdGripOpen);
_rtrigGripClose(CLK := _bCmdGripClose);

(* Safety edge detection from safe output byte 0 *)
_rtrigSafeStop1(CLK := _bSafeCmdSS1);
_rtrigSafeEStop(CLK := _bSafeCmdEStop);

(* Requested job number: bytes 2-3 WORD LE, or byte 2 only (GVL_Program.JOB_NUMBER_BYTE) *)
IF GVL_Program.JOB_NUMBER_BYTE THEN
    _wRequestedJob := BYTE_TO_WORD(aVassOutputData[2]);
ELSE
    _wRequestedJob := BYTE_TO_WORD(aVassOutputData[2])
                      OR SHL(BYTE_TO_WORD(aVassOutputData[3]), 8);
END_IF

(* Zone GRANT: DWORD LE at bytes GVL_Program.GRANT_BYTE..+3 *)
_nIdx := GVL_Program.GRANT_BYTE;
_dwGrant := BYTE_TO_DWORD(aVassOutputData[_nIdx])
            OR SHL(BYTE_TO_DWORD(aVassOutputData[_nIdx + 1]), 8)
            OR SHL(BYTE_TO_DWORD(aVassOutputData[_nIdx + 2]), 16)
            OR SHL(BYTE_TO_DWORD(aVassOutputData[_nIdx + 3]), 24);

(* ============================================================================
   SECTION 2: SAFETY LOGIC (PROFIsafe Slot 1)
   Reads abySafeOut, status is written to abySafeIn in section 4
   ============================================================================ *)

(* Process safe outputs from PLC - byte 0 *)
_bSafe_DrivesOK := _bSafeCmdDriveEnable AND _bSafe_EStopOK AND NOT _bSafe_Fault;

(* E-Stop handling *)
IF _bSafeCmdEStop THEN  (* External E-Stop *)
    _bSafe_EStopOK := FALSE;
    _bSafe_STO := TRUE;
    _bDrivesPowered := FALSE;
    _bProgRunning := FALSE;
    eProgramState := E_ProgramState#PRG_STOPPED;
END_IF

(* Safe Stop 1 request *)
IF _bSafeCmdSS1 AND _bProgRunning THEN
    _bSafe_SS1 := TRUE;
    _bProgRunning := FALSE;
    _bSafe_Stopped := TRUE;
    eProgramState := E_ProgramState#PRG_STOPPED;
END_IF

(* Recovery from safety state *)
IF NOT _bSafeCmdEStop AND NOT _bSafeCmdSS1 THEN
    IF _bCmdReset THEN  (* Reset bit *)
        _bSafe_EStopOK := TRUE;
        _bSafe_STO := FALSE;
        _bSafe_SS1 := FALSE;
        _bSafe_Stopped := FALSE;
        _bSafe_Fault := FALSE;
    END_IF
END_IF

(* Overall safety status *)
bSafetyOK := _bSafe_DrivesOK AND _bSafe_EStopOK AND _bSafe_GatesClosed AND NOT _bSafe_Fault;
_bSafe_GatesClosed := TRUE; (* Always closed in simulation *)

(* ============================================================================
   SECTION 3: STANDARD I/O LOGIC (VASS Telegram Slot 2)
   ============================================================================ *)

(* --- Drive Power Control --- *)
_tonDriveStartup(IN := _bCmdDrivesOn AND bSafetyOK AND NOT _bDrivesPowered, PT := T#2S);
IF _tonDriveStartup.Q THEN
    _bDrivesPowered := TRUE;
    _bSafe_Stopped := FALSE;
END_IF

IF NOT _bCmdDrivesOn OR NOT bSafetyOK THEN
    _bDrivesPowered := FALSE;
    _bProgRunning := FALSE;
    IF eProgramState = E_ProgramState#PRG_RUNNING THEN
        eProgramState := E_ProgramState#PRG_STOPPED;
    END_IF
END_IF

(* --- Mode Control --- *)
_bInExtMode := _bCmdModeExt AND _bDrivesPowered AND bSafetyOK;
IF _bInExtMode THEN
    eCurrentMode := E_RobotMode#MODE_EXT;
ELSE
    eCurrentMode := E_RobotMode#MODE_T1;
END_IF

(* --- Ready State --- *)
_bReady := _bDrivesPowered
           AND _bInExtMode
           AND NOT _bError
           AND NOT _bProgRunning
           AND bSafetyOK;

(* --- Warning reset: any Reset edge clears a pending warning (no error needed) --- *)
IF _rtrigReset.Q THEN
    _wWarningCode := WORD#0;
END_IF

(* --- Error Reset (Reset held 500 ms) --- *)
_tonErrorReset(IN := _bCmdReset AND _bError, PT := T#500MS);
IF _tonErrorReset.Q THEN
    _bError := FALSE;
    _wErrorCode := WORD#0;
    _wWarningCode := WORD#0;
    IF eProgramState = E_ProgramState#PRG_ERROR THEN
        eProgramState := E_ProgramState#PRG_IDLE;
    END_IF
END_IF

(* --- Job Request Handling --- *)
IF _rtrigJobReq.Q AND _bReady THEN
    _wActiveJob := _wRequestedJob;
    _bJobAcknowledged := TRUE;
    _bProgFinished := FALSE;
    (* PLAN_ID: WORD LE at bytes GVL_Program.PLAN_ID_BYTE..+1 (production job only) *)
    _nIdx := GVL_Program.PLAN_ID_BYTE;
    _wPlanId := BYTE_TO_WORD(aVassOutputData[_nIdx])
                OR SHL(BYTE_TO_WORD(aVassOutputData[_nIdx + 1]), 8);
END_IF

IF NOT _bCmdJobReq THEN
    _bJobAcknowledged := FALSE;
END_IF

(* --- Program Start --- *)
_bStartOk := FALSE;
IF _rtrigProgStart.Q AND _bReady AND _wActiveJob <> WORD#0 THEN
    _wPlayerJob := _wActiveJob;
    IF _wActiveJob = GVL_Program.HOME_FOLGE THEN
        _bStartOk := TRUE;
    ELSIF _wActiveJob = GVL_Program.PROD_FOLGE AND GVL_Program.N_OPS > 0 THEN
        IF _wPlanId = GVL_Program.PLAN_ID THEN
            _bStartOk := TRUE;
        ELSE
            _bError := TRUE;
            _wErrorCode := GVL_Program.ERR_PLAN_MISMATCH;
            eProgramState := E_ProgramState#PRG_ERROR;
        END_IF
    ELSE
        _bError := TRUE;
        _wErrorCode := GVL_Program.ERR_UNKNOWN_FOLGE;
        eProgramState := E_ProgramState#PRG_ERROR;
    END_IF
ELSIF _rtrigHome.Q AND _bReady AND NOT _bAtHome THEN
    (* HomeRequest [0].6 edge while Ready: behaves like HOME_FOLGE *)
    _wPlayerJob := GVL_Program.HOME_FOLGE;
    _bStartOk := TRUE;
END_IF

IF _bStartOk THEN
    _bProgRunning := TRUE;
    _bProgFinished := FALSE;
    _bInPosition := FALSE;
    _bSafe_Stopped := FALSE;
    _bPlayerStart := TRUE;
    eProgramState := E_ProgramState#PRG_RUNNING;
END_IF

(* --- Program Stop/Cancel (level) --- *)
IF (_bCmdProgStop OR _bCmdProgCancel) AND _bProgRunning THEN
    _bProgRunning := FALSE;
    _bProgFinished := FALSE;
    _bInPosition := TRUE;
    eProgramState := E_ProgramState#PRG_STOPPED;
END_IF

(* --- Program Execution: FB_ProgramPlayer --- *)
(* Any stop path above (Stop/Cancel, drives off, E-stop, SS1) aborts the player in this scan:
   REQUEST := 0, step := 0, the pose is held. *)
_rRate := UINT_TO_REAL(WORD_TO_UINT(_wSpeed)) / 100.0;
_fbPlayer(
    bStart  := _bPlayerStart,
    wJob    := _wPlayerJob,
    bAbort  := NOT _bProgRunning,
    dwGrant := _dwGrant,
    rRate   := _rRate,
    rDt     := rDt
);
_bPlayerStart := FALSE;

IF _bProgRunning THEN
    IF _fbPlayer.bError THEN
        _bProgRunning := FALSE;
        _bError := TRUE;
        _wErrorCode := _fbPlayer.wErrorCode;
        eProgramState := E_ProgramState#PRG_ERROR;
    ELSIF _fbPlayer.bDone THEN
        (* Same scan as step := 0: ProgRunning drops and ProgFinished rises together *)
        _bProgRunning := FALSE;
        _bProgFinished := TRUE;
        _bInPosition := TRUE;
        eProgramState := E_ProgramState#PRG_FINISHED;
    END_IF
END_IF

_wCurrentStep := _fbPlayer.wStep;
_dwRequest := _fbPlayer.dwRequest;
_bAtHome := _fbPlayer.bAtHome;

(* Player warnings are copied on change, so an error reset clears them *)
IF _fbPlayer.wWarningCode <> _wPlayerWarning THEN
    _wPlayerWarning := _fbPlayer.wWarningCode;
    IF _wPlayerWarning <> WORD#0 THEN
        _wWarningCode := _wPlayerWarning;
    END_IF
END_IF

(* --- Gripper Simulation --- *)
_tonGripperAction(IN := _bCmdGripClose AND NOT _bGripperClosed, PT := T#500MS);
IF _tonGripperAction.Q THEN
    _bGripperClosed := TRUE;
    _bPartPresent := TRUE;
END_IF

IF _bCmdGripOpen THEN
    _bGripperClosed := FALSE;
    _bPartPresent := FALSE;
END_IF

(* --- Speed Override (bytes 8-9 WORD LE, applied with [1].4) --- *)
_wSpeedCmd := BYTE_TO_WORD(aVassOutputData[8]) OR SHL(BYTE_TO_WORD(aVassOutputData[9]), 8);
IF _bCmdSpeedOverride AND WORD_TO_UINT(_wSpeedCmd) > 0 AND WORD_TO_UINT(_wSpeedCmd) <= 100 THEN
    _wSpeed := _wSpeedCmd;
END_IF

(* ============================================================================
   SECTION 4: WRITE SAFETY STATUS to abySafeIn[0..7]
   ============================================================================ *)

(* Byte 0: Safe drive/motion status *)
abySafeIn[0].0 := _bSafe_DrivesOK;
abySafeIn[0].1 := _bSafe_Stopped;
abySafeIn[0].2 := FALSE; (* Reduced speed *)
abySafeIn[0].3 := NOT _bSafe_Fault; (* Axis monitor OK *)
abySafeIn[0].4 := TRUE;  (* Tool monitor OK *)
abySafeIn[0].5 := TRUE;  (* Workspace OK *)
abySafeIn[0].6 := FALSE;
abySafeIn[0].7 := FALSE;

(* Byte 1: Gate/protection status *)
abySafeIn[1].0 := _bSafe_GatesClosed;  (* Gate 1 *)
abySafeIn[1].1 := _bSafe_GatesClosed;  (* Gate 2 *)
abySafeIn[1].2 := _bSafe_GatesClosed;  (* Gate 3 *)
abySafeIn[1].3 := TRUE;   (* Light curtain OK *)
abySafeIn[1].4 := _bSafe_EStopOK;
abySafeIn[1].5 := FALSE;  (* Enabling device *)
abySafeIn[1].6 := TRUE;   (* Operator safe *)
abySafeIn[1].7 := FALSE;

(* Byte 2: Extended safe functions *)
abySafeIn[2].0 := _bSafe_STO;
abySafeIn[2].1 := _bSafe_SS1;
abySafeIn[2].2 := FALSE;  (* SS2 *)
abySafeIn[2].3 := _bSafe_Stopped AND NOT _bSafe_STO;  (* SOS *)
abySafeIn[2].4 := FALSE;  (* SLS *)
abySafeIn[2].5 := FALSE;  (* SLP *)
abySafeIn[2].6 := FALSE;
abySafeIn[2].7 := _bSafe_Fault;

(* Bytes 3-7: zero *)
abySafeIn[3] := BYTE#0;
abySafeIn[4] := BYTE#0;
abySafeIn[5] := BYTE#0;
abySafeIn[6] := BYTE#0;
abySafeIn[7] := BYTE#0;

(* ============================================================================
   SECTION 5: WRITE VASS STATUS to aVassInputData[0..31]
   ============================================================================ *)

(* Unused bytes are zero; bytes 16-27 (joint angles) are filled by PLC_PRG *)
FOR _i := 0 TO 31 DO
    aVassInputData[_i] := BYTE#0;
END_FOR

(* Status Word - Byte 0 *)
aVassInputData[0].0 := _bDrivesPowered;
aVassInputData[0].1 := _bProgRunning;
aVassInputData[0].2 := _bAtHome;
aVassInputData[0].3 := _bInPosition;
aVassInputData[0].4 := _bInExtMode;
aVassInputData[0].5 := _bReady;
aVassInputData[0].6 := _bError;
aVassInputData[0].7 := _wWarningCode <> WORD#0;

(* Status Word - Byte 1 *)
aVassInputData[1].0 := _bSafe_GatesClosed;
aVassInputData[1].1 := _bSafe_EStopOK;
aVassInputData[1].2 := _bProgFinished;
aVassInputData[1].3 := _bJobAcknowledged;
aVassInputData[1].4 := _bGripperClosed;
aVassInputData[1].5 := _bPartPresent;
aVassInputData[1].6 := TRUE;  (* Periph ready *)
aVassInputData[1].7 := FALSE; (* Maint not required *)

(* Active job number echo - Bytes 2-3 (byte 2 only in byte mode, byte 3 = 0) *)
aVassInputData[2] := WORD_TO_BYTE(_wActiveJob AND WORD#16#FF);
IF NOT GVL_Program.JOB_NUMBER_BYTE THEN
    aVassInputData[3] := WORD_TO_BYTE(SHR(_wActiveJob, 8));
END_IF

(* Speed actual - Bytes 6-7 *)
aVassInputData[6] := WORD_TO_BYTE(_wSpeed AND WORD#16#FF);
aVassInputData[7] := WORD_TO_BYTE(SHR(_wSpeed, 8));

(* Tool number - Bytes 8-9 *)
aVassInputData[8] := WORD_TO_BYTE(_wToolNr AND WORD#16#FF);
aVassInputData[9] := WORD_TO_BYTE(SHR(_wToolNr, 8));

(* Error code - Bytes 10-11 *)
aVassInputData[10] := WORD_TO_BYTE(_wErrorCode AND WORD#16#FF);
aVassInputData[11] := WORD_TO_BYTE(SHR(_wErrorCode, 8));

(* Warning code - Bytes 12-13 *)
aVassInputData[12] := WORD_TO_BYTE(_wWarningCode AND WORD#16#FF);
aVassInputData[13] := WORD_TO_BYTE(SHR(_wWarningCode, 8));

(* Position X - Bytes 14-15 *)
aVassInputData[14] := WORD_TO_BYTE(INT_TO_WORD(_iPositionX) AND WORD#16#FF);
aVassInputData[15] := WORD_TO_BYTE(SHR(INT_TO_WORD(_iPositionX), 8));

(* Bytes 16-27: A129_224_Option area - RESERVED for the joint angle encoder
   (PLC_PRG -> fbJointEncoder, 6x INT big-endian = A1..A6 at 0.02 deg/count) *)

(* Current step (op index) - WORD LE at bytes GVL_Program.STEP_BYTE..+1 *)
_nIdx := GVL_Program.STEP_BYTE;
aVassInputData[_nIdx] := WORD_TO_BYTE(_wCurrentStep AND WORD#16#FF);
aVassInputData[_nIdx + 1] := WORD_TO_BYTE(SHR(_wCurrentStep, 8));

(* Zone REQUEST - DWORD LE at bytes GVL_Program.REQ_BYTE..+3 *)
_nIdx := GVL_Program.REQ_BYTE;
aVassInputData[_nIdx] := DWORD_TO_BYTE(_dwRequest AND DWORD#16#FF);
aVassInputData[_nIdx + 1] := DWORD_TO_BYTE(SHR(_dwRequest, 8) AND DWORD#16#FF);
aVassInputData[_nIdx + 2] := DWORD_TO_BYTE(SHR(_dwRequest, 16) AND DWORD#16#FF);
aVassInputData[_nIdx + 3] := DWORD_TO_BYTE(SHR(_dwRequest, 24));

(* ============================================================================
   SECTION 6: OUTPUTS (joint angles, diagnostics)
   ============================================================================ *)
rA1_deg := _fbPlayer.rA1_deg;
rA2_deg := _fbPlayer.rA2_deg;
rA3_deg := _fbPlayer.rA3_deg;
rA4_deg := _fbPlayer.rA4_deg;
rA5_deg := _fbPlayer.rA5_deg;
rA6_deg := _fbPlayer.rA6_deg;

wActiveJob := _wActiveJob;
wCurrentStep := _wCurrentStep;
wErrorCode := _wErrorCode;
dwRequest := _dwRequest;
dwGrant := _dwGrant;
ePlayerState := _fbPlayer.eState;
END_FUNCTION_BLOCK
